Universal Robots URScript: FaiChun_9 Jan_Mcam1.script

def Machining1():
  # Default parameters:
  global speed_ms = 0.05
  global speed_rads = 0.75
  global accel_mss = 3
  global accel_radss = 1.2
  global blend_radius_m = 0.0003

  # Add subprograms here
  # Start of main program
  # Program generated by RoboDK v5.6.8 for UR10e on 13/01/2025 15:21:15
  # Using nominal kinematics.
  blend_radius_m = 0.0003
  speed_ms = 0.05
  # set_reference(p[0.340000, -0.055000, 0.001500, 0.000000, 0.000000, 0.000000])
  set_tcp(p[0.000000, 0.000000, 0.252000, 0.000000, 0.000000, 0.000000])
  # Show Tool
  movej([0.369740, -1.015857, -2.630541, -1.065992, 1.570796, 1.940536],accel_radss,speed_rads,0,blend_radius_m)
  movel([0.369740, -1.070501, -2.672301, -0.969586, 1.570796, 1.940536],accel_mss,speed_ms,0,blend_radius_m)
  #SetTool218
  #M_RunCode6
  #SetRPM107900
  #M_RunCode3
  speed_ms = 0.05
  movel([0.369740, -1.102928, -2.692299, -0.917162, 1.570796, 1.940536],accel_mss,speed_ms,0,blend_radius_m)
  speed_ms = 0.017
  movel([0.369740, -1.139169, -2.711618, -0.861603, 1.570796, 1.940536],accel_mss,speed_ms,0,blend_radius_m)
  speed_ms = 0.051
  movel([0.740413, -1.151810, -2.706369, -0.854210, 1.570796, 2.311209],accel_mss,speed_ms,0,blend_radius_m)
  movel([0.532956, -1.474706, -2.506843, -0.730840, 1.570796, 2.103752],accel_mss,speed_ms,0,blend_radius_m)
  movel([0.260506, -1.469805, -2.510970, -0.731614, 1.570796, 1.831302],accel_mss,speed_ms,0,blend_radius_m)
  movel([0.369740, -1.139169, -2.711618, -0.861603, 1.570796, 1.940536],accel_mss,speed_ms,0,blend_radius_m)
  speed_ms = 0.05
  movel([0.369740, -1.070501, -2.672301, -0.969586, 1.570796, 1.940536],accel_mss,speed_ms,0,blend_radius_m)
  speed_ms = 0.051
  movel([0.403329, -1.072947, -2.671379, -0.968064, 1.570796, 1.974125],accel_mss,speed_ms,0,blend_radius_m)
  movel([0.403329, -1.105379, -2.691338, -0.915672, 1.570796, 1.974125],accel_mss,speed_ms,0,blend_radius_m)
  speed_ms = 0.017
  movel([0.403329, -1.141610, -2.710617, -0.860163, 1.570796, 1.974125],accel_mss,speed_ms,0,blend_radius_m)
  speed_ms = 0.051
  movel([0.704795, -1.151689, -2.706421, -0.854280, 1.570796, 2.275591],accel_mss,speed_ms,0,blend_radius_m)
  movel([0.696497, -1.164526, -2.700927, -0.846935, 1.570796, 2.267294],accel_mss,speed_ms,0,blend_radius_m)
  movel([0.703914, -1.166306, -2.700152, -0.845930, 1.570796, 2.274710],accel_mss,speed_ms,0,blend_radius_m)
  movel([0.706062, -1.163020, -2.701581, -0.847789, 1.570796, 2.276858],accel_mss,speed_ms,0,blend_radius_m)
  movel([0.701176, -1.161829, -2.702095, -0.848464, 1.570796, 2.271972],accel_mss,speed_ms,0,blend_radius_m)
  movel([0.707357, -1.152320, -2.706154, -0.853914, 1.570796, 2.278154],accel_mss,speed_ms,0,blend_radius_m)
  movel([0.714620, -1.154134, -2.705387, -0.852868, 1.570796, 2.285416],accel_mss,speed_ms,0,blend_radius_m)
  movel([0.710409, -1.160546, -2.702649, -0.849195, 1.570796, 2.281205],accel_mss,speed_ms,0,blend_radius_m)
  movel([0.712930, -1.161189, -2.702372, -0.848829, 1.570796, 2.283727],accel_mss,speed_ms,0,blend_radius_m)
  movel([0.717151, -1.154792, -2.705108, -0.852489, 1.570796, 2.287947],accel_mss,speed_ms,0,blend_radius_m)
  movel([0.724331, -1.156706, -2.704294, -0.851389, 1.570796, 2.295128],accel_mss,speed_ms,0,blend_radius_m)
  movel([0.720088, -1.163073, -2.701558, -0.847759, 1.570796, 2.290884],accel_mss,speed_ms,0,blend_radius_m)
  movel([0.724885, -1.164384, -2.700989, -0.847016, 1.570796, 2.295682],accel_mss,speed_ms,0,blend_radius_m)
  movel([0.718665, -1.173659, -2.696916, -0.841814, 1.570796, 2.289462],accel_mss,speed_ms,0,blend_radius_m)
  movel([0.713893, -1.172379, -2.697484, -0.842526, 1.570796, 2.284689],accel_mss,speed_ms,0,blend_radius_m)
  movel([0.711746, -1.175609, -2.696048, -0.840731, 1.570796, 2.282542],accel_mss,speed_ms,0,blend_radius_m)
  movel([0.716510, -1.176879, -2.695481, -0.840029, 1.570796, 2.287306],accel_mss,speed_ms,0,blend_radius_m)
  movel([0.710435, -1.185964, -2.691373, -0.835052, 1.570796, 2.281231],accel_mss,speed_ms,0,blend_radius_m)
  movel([0.703407, -1.184139, -2.692206, -0.836045, 1.570796, 2.274203],accel_mss,speed_ms,0,blend_radius_m)
  movel([0.707472, -1.177990, -2.694983, -0.839416, 1.570796, 2.278268],accel_mss,speed_ms,0,blend_radius_m)
  movel([0.704985, -1.177355, -2.695268, -0.839766, 1.570796, 2.275781],accel_mss,speed_ms,0,blend_radius_m)
  movel([0.698841, -1.186688, -2.691042, -0.834659, 1.570796, 2.269637],accel_mss,speed_ms,0,blend_radius_m)
  movel([0.708330, -1.189119, -2.689926, -0.833344, 1.570796, 2.279126],accel_mss,speed_ms,0,blend_radius_m)
  movel([0.541731, -1.451056, -2.526411, -0.734922, 1.570796, 2.112528],accel_mss,speed_ms,0,blend_radius_m)
  movel([0.533908, -1.449838, -2.527395, -0.735156, 1.570796, 2.104704],accel_mss,speed_ms,0,blend_radius_m)
  movel([0.530407, -1.455837, -2.522525, -0.734027, 1.570796, 2.101203],accel_mss,speed_ms,0,blend_radius_m)
  movel([0.532431, -1.456143, -2.522276, -0.733971, 1.570796, 2.103227],accel_mss,speed_ms,0,blend_radius_m)
  movel([0.534734, -1.452207, -2.525478, -0.734704, 1.570796, 2.105531],accel_mss,speed_ms,0,blend_radius_m)
  movel([0.540507, -1.453110, -2.524746, -0.734533, 1.570796, 2.111303],accel_mss,speed_ms,0,blend_radius_m)
  movel([0.537071, -1.458916, -2.520004, -0.733469, 1.570796, 2.107867],accel_mss,speed_ms,0,blend_radius_m)
  movel([0.533196, -1.458312, -2.520500, -0.733577, 1.570796, 2.103992],accel_mss,speed_ms,0,blend_radius_m)
  movel([0.532009, -1.460340, -2.518833, -0.733216, 1.570796, 2.102805],accel_mss,speed_ms,0,blend_radius_m)
  movel([0.535879, -1.460941, -2.518338, -0.733110, 1.570796, 2.106675],accel_mss,speed_ms,0,blend_radius_m)
  movel([0.532503, -1.466680, -2.513581, -0.732128, 1.570796, 2.103300],accel_mss,speed_ms,0,blend_radius_m)
  movel([0.528655, -1.466088, -2.514074, -0.732226, 1.570796, 2.099451],accel_mss,speed_ms,0,blend_radius_m)
  movel([0.526411, -1.469942, -2.510855, -0.731592, 1.570796, 2.097208],accel_mss,speed_ms,0,blend_radius_m)
  movel([0.520712, -1.469102, -2.511559, -0.731728, 1.570796, 2.091509],accel_mss,speed_ms,0,blend_radius_m)
  movel([0.522933, -1.465238, -2.514782, -0.732370, 1.570796, 2.093730],accel_mss,speed_ms,0,blend_radius_m)
  movel([0.520922, -1.464950, -2.515020, -0.732418, 1.570796, 2.091718],accel_mss,speed_ms,0,blend_radius_m)
  movel([0.518707, -1.468815, -2.511798, -0.731775, 1.570796, 2.089503],accel_mss,speed_ms,0,blend_radius_m)
  movel([0.512973, -1.468021, -2.512463, -0.731905, 1.570796, 2.083769],accel_mss,speed_ms,0,blend_radius_m)
  movel([0.516230, -1.462277, -2.517236, -0.732877, 1.570796, 2.087027],accel_mss,speed_ms,0,blend_radius_m)
  movel([0.520125, -1.462817, -2.516788, -0.732783, 1.570796, 2.090921],accel_mss,speed_ms,0,blend_radius_m)
  movel([0.521283, -1.460796, -2.518457, -0.733135, 1.570796, 2.092080],accel_mss,speed_ms,0,blend_radius_m)
  movel([0.515352, -1.459974, -2.519134, -0.733281, 1.570796, 2.086148],accel_mss,speed_ms,0,blend_radius_m)
  movel([0.510955, -1.467752, -2.512687, -0.731950, 1.570796, 2.081751],accel_mss,speed_ms,0,blend_radius_m)
  movel([0.287607, -1.463384, -2.516319, -0.732685, 1.570796, 1.858403],accel_mss,speed_ms,0,blend_radius_m)
  movel([0.290165, -1.455515, -2.522788, -0.734086, 1.570796, 1.860961],accel_mss,speed_ms,0,blend_radius_m)
  movel([0.283577, -1.456094, -2.522316, -0.733980, 1.570796, 1.854374],accel_mss,speed_ms,0,blend_radius_m)
  movel([0.282922, -1.458141, -2.520640, -0.733608, 1.570796, 1.853718],accel_mss,speed_ms,0,blend_radius_m)
  movel([0.287251, -1.457756, -2.520955, -0.733677, 1.570796, 1.858048],accel_mss,speed_ms,0,blend_radius_m)
  movel([0.285369, -1.463569, -2.516166, -0.732654, 1.570796, 1.856165],accel_mss,speed_ms,0,blend_radius_m)
  movel([0.279002, -1.464133, -2.515698, -0.732557, 1.570796, 1.849799],accel_mss,speed_ms,0,blend_radius_m)
  movel([0.280240, -1.460222, -2.518931, -0.733237, 1.570796, 1.851036],accel_mss,speed_ms,0,blend_radius_m)
  movel([0.277998, -1.460430, -2.518759, -0.733200, 1.570796, 1.848794],accel_mss,speed_ms,0,blend_radius_m)
  movel([0.276770, -1.464340, -2.515527, -0.732522, 1.570796, 1.847566],accel_mss,speed_ms,0,blend_radius_m)
  movel([0.270394, -1.464949, -2.515021, -0.732418, 1.570796, 1.841191],accel_mss,speed_ms,0,blend_radius_m)
  movel([0.271594, -1.461046, -2.518252, -0.733092, 1.570796, 1.842390],accel_mss,speed_ms,0,blend_radius_m)
  movel([0.267266, -1.461483, -2.517891, -0.733015, 1.570796, 1.838062],accel_mss,speed_ms,0,blend_radius_m)
  movel([0.269033, -1.455666, -2.522665, -0.734058, 1.570796, 1.839830],accel_mss,speed_ms,0,blend_radius_m)
  movel([0.273388, -1.455222, -2.523027, -0.734140, 1.570796, 1.844184],accel_mss,speed_ms,0,blend_radius_m)
  movel([0.274023, -1.453169, -2.524697, -0.734522, 1.570796, 1.844820],accel_mss,speed_ms,0,blend_radius_m)
  movel([0.269656, -1.453615, -2.524335, -0.734439, 1.570796, 1.840452],accel_mss,speed_ms,0,blend_radius_m)
  movel([0.271457, -1.447728, -2.529094, -0.735567, 1.570796, 1.842253],accel_mss,speed_ms,0,blend_radius_m)
  movel([0.277970, -1.447061, -2.529630, -0.735698, 1.570796, 1.848766],accel_mss,speed_ms,0,blend_radius_m)
  movel([0.276719, -1.451051, -2.526415, -0.734923, 1.570796, 1.847516],accel_mss,speed_ms,0,blend_radius_m)
  movel([0.278991, -1.450829, -2.526594, -0.734966, 1.570796, 1.849787],accel_mss,speed_ms,0,blend_radius_m)
  movel([0.280907, -1.444757, -2.531476, -0.736156, 1.570796, 1.851704],accel_mss,speed_ms,0,blend_radius_m)
  movel([0.272096, -1.445651, -2.530761, -0.735977, 1.570796, 1.842893],accel_mss,speed_ms,0,blend_radius_m)
  movel([0.361539, -1.178261, -2.694862, -0.839266, 1.570796, 1.932335],accel_mss,speed_ms,0,blend_radius_m)
  movel([0.373305, -1.176443, -2.695676, -0.840270, 1.570796, 1.944101],accel_mss,speed_ms,0,blend_radius_m)
  movel([0.376834, -1.166854, -2.699913, -0.845622, 1.570796, 1.947630],accel_mss,speed_ms,0,blend_radius_m)
  movel([0.373758, -1.167323, -2.699708, -0.845358, 1.570796, 1.944554],accel_mss,speed_ms,0,blend_radius_m)
  movel([0.371445, -1.173642, -2.696924, -0.841824, 1.570796, 1.942241],accel_mss,speed_ms,0,blend_radius_m)
  movel([0.362714, -1.175005, -2.696318, -0.841066, 1.570796, 1.933510],accel_mss,speed_ms,0,blend_radius_m)
  movel([0.366061, -1.165657, -2.700435, -0.846297, 1.570796, 1.936857],accel_mss,speed_ms,0,blend_radius_m)
  movel([0.372018, -1.164705, -2.700850, -0.846834, 1.570796, 1.942815],accel_mss,speed_ms,0,blend_radius_m)
  movel([0.373227, -1.161386, -2.702286, -0.848716, 1.570796, 1.944024],accel_mss,speed_ms,0,blend_radius_m)
  movel([0.367253, -1.162346, -2.701872, -0.848171, 1.570796, 1.938049],accel_mss,speed_ms,0,blend_radius_m)
  movel([0.370690, -1.152795, -2.705954, -0.853640, 1.570796, 1.941486],accel_mss,speed_ms,0,blend_radius_m)
  movel([0.376724, -1.151811, -2.706369, -0.854209, 1.570796, 1.947521],accel_mss,speed_ms,0,blend_radius_m)
  movel([0.379122, -1.145259, -2.709109, -0.858021, 1.570796, 1.949918],accel_mss,speed_ms,0,blend_radius_m)
  movel([0.388102, -1.143842, -2.709696, -0.858851, 1.570796, 1.958898],accel_mss,speed_ms,0,blend_radius_m)
  movel([0.385643, -1.150419, -2.706955, -0.855015, 1.570796, 1.956439],accel_mss,speed_ms,0,blend_radius_m)
  movel([0.388764, -1.149949, -2.707152, -0.855288, 1.570796, 1.959560],accel_mss,speed_ms,0,blend_radius_m)
  movel([0.391247, -1.143361, -2.709895, -0.859133, 1.570796, 1.962043],accel_mss,speed_ms,0,blend_radius_m)
  movel([0.400196, -1.142054, -2.710434, -0.859901, 1.570796, 1.970993],accel_mss,speed_ms,0,blend_radius_m)
  movel([0.396453, -1.151808, -2.706370, -0.854211, 1.570796, 1.967249],accel_mss,speed_ms,0,blend_radius_m)
  movel([0.390466, -1.152664, -2.706009, -0.853716, 1.570796, 1.961262],accel_mss,speed_ms,0,blend_radius_m)
  movel([0.389190, -1.156041, -2.704577, -0.851771, 1.570796, 1.959986],accel_mss,speed_ms,0,blend_radius_m)
  movel([0.398252, -1.154767, -2.705119, -0.852504, 1.570796, 1.969048],accel_mss,speed_ms,0,blend_radius_m)
  movel([0.403329, -1.141610, -2.710617, -0.860163, 1.570796, 1.974125],accel_mss,speed_ms,0,blend_radius_m)
  speed_ms = 0.05
  movel([0.403329, -1.072947, -2.671379, -0.968064, 1.570796, 1.974125],accel_mss,speed_ms,0,blend_radius_m)
  #M_RunCode5
  speed_ms = 0.051
  movel([0.436039, -1.030309, -2.635411, -1.046670, 1.570796, 2.006835],accel_mss,speed_ms,0,blend_radius_m)
  #M_RunCode1
  #SetTool213
  #M_RunCode6
  #SetRPM107900
  #M_RunCode3
  speed_ms = 0.05
  movel([0.380621, -0.927251, -2.391546, -1.393592, 1.570796, 1.951417],accel_mss,speed_ms,0,blend_radius_m)
  speed_ms = 0.051
  movel([0.380621, -1.121069, -2.652122, -0.939198, 1.570796, 1.951417],accel_mss,speed_ms,0,blend_radius_m)
  movel([0.380621, -1.153481, -2.671325, -0.887584, 1.570796, 1.951417],accel_mss,speed_ms,0,blend_radius_m)
  speed_ms = 0.017
  movel([0.380621, -1.189377, -2.689807, -0.833205, 1.570796, 1.951417],accel_mss,speed_ms,0,blend_radius_m)
  speed_ms = 0.051
  movel([0.383999, -1.188172, -2.690361, -0.833856, 1.570796, 1.954796],accel_mss,speed_ms,0,blend_radius_m)
  movel([0.387929, -1.187302, -2.690760, -0.834326, 1.570796, 1.958725],accel_mss,speed_ms,0,blend_radius_m)
  movel([0.392921, -1.186724, -2.691025, -0.834640, 1.570796, 1.963717],accel_mss,speed_ms,0,blend_radius_m)
  movel([0.396406, -1.186468, -2.691143, -0.834778, 1.570796, 1.967202],accel_mss,speed_ms,0,blend_radius_m)
  movel([0.399894, -1.186176, -2.691276, -0.834937, 1.570796, 1.970690],accel_mss,speed_ms,0,blend_radius_m)
  movel([0.403055, -1.185763, -2.691465, -0.835161, 1.570796, 1.973851],accel_mss,speed_ms,0,blend_radius_m)
  movel([0.405472, -1.185291, -2.691681, -0.835418, 1.570796, 1.976268],accel_mss,speed_ms,0,blend_radius_m)
  movel([0.407571, -1.184727, -2.691938, -0.835724, 1.570796, 1.978367],accel_mss,speed_ms,0,blend_radius_m)
  movel([0.410903, -1.183473, -2.692508, -0.836408, 1.570796, 1.981699],accel_mss,speed_ms,0,blend_radius_m)
  movel([0.412588, -1.182637, -2.692888, -0.836864, 1.570796, 1.983384],accel_mss,speed_ms,0,blend_radius_m)
  movel([0.415576, -1.180774, -2.693730, -0.837884, 1.570796, 1.986373],accel_mss,speed_ms,0,blend_radius_m)
  movel([0.417237, -1.179418, -2.694342, -0.838629, 1.570796, 1.988033],accel_mss,speed_ms,0,blend_radius_m)
  movel([0.418646, -1.177700, -2.695113, -0.839575, 1.570796, 1.989443],accel_mss,speed_ms,0,blend_radius_m)
  movel([0.419750, -1.175666, -2.696023, -0.840700, 1.570796, 1.990546],accel_mss,speed_ms,0,blend_radius_m)
  movel([0.420402, -1.173479, -2.696996, -0.841914, 1.570796, 1.991198],accel_mss,speed_ms,0,blend_radius_m)
  movel([0.420438, -1.171501, -2.697872, -0.843016, 1.570796, 1.991235],accel_mss,speed_ms,0,blend_radius_m)
  movel([0.420217, -1.170743, -2.698207, -0.843440, 1.570796, 1.991013],accel_mss,speed_ms,0,blend_radius_m)
  movel([0.419855, -1.170173, -2.698457, -0.843759, 1.570796, 1.990652],accel_mss,speed_ms,0,blend_radius_m)
  movel([0.419383, -1.169789, -2.698626, -0.843973, 1.570796, 1.990180],accel_mss,speed_ms,0,blend_radius_m)
  movel([0.418119, -1.169559, -2.698728, -0.844102, 1.570796, 1.988915],accel_mss,speed_ms,0,blend_radius_m)
  movel([0.416505, -1.170034, -2.698519, -0.843836, 1.570796, 1.987302],accel_mss,speed_ms,0,blend_radius_m)
  movel([0.416237, -1.170163, -2.698462, -0.843764, 1.570796, 1.987034],accel_mss,speed_ms,0,blend_radius_m)
  movel([0.414985, -1.171929, -2.697683, -0.842778, 1.570796, 1.985782],accel_mss,speed_ms,0,blend_radius_m)
  movel([0.413492, -1.173744, -2.696878, -0.841766, 1.570796, 1.984288],accel_mss,speed_ms,0,blend_radius_m)
  movel([0.412436, -1.174807, -2.696406, -0.841176, 1.570796, 1.983232],accel_mss,speed_ms,0,blend_radius_m)
  movel([0.411578, -1.175521, -2.696088, -0.840780, 1.570796, 1.982374],accel_mss,speed_ms,0,blend_radius_m)
  movel([0.410708, -1.176097, -2.695830, -0.840461, 1.570796, 1.981504],accel_mss,speed_ms,0,blend_radius_m)
  movel([0.409905, -1.176478, -2.695660, -0.840250, 1.570796, 1.980701],accel_mss,speed_ms,0,blend_radius_m)
  movel([0.408376, -1.176754, -2.695537, -0.840098, 1.570796, 1.979172],accel_mss,speed_ms,0,blend_radius_m)
  movel([0.408234, -1.176742, -2.695542, -0.840104, 1.570796, 1.979030],accel_mss,speed_ms,0,blend_radius_m)
  movel([0.406466, -1.176296, -2.695742, -0.840351, 1.570796, 1.977262],accel_mss,speed_ms,0,blend_radius_m)
  movel([0.405390, -1.175348, -2.696165, -0.840876, 1.570796, 1.976186],accel_mss,speed_ms,0,blend_radius_m)
  movel([0.404939, -1.173986, -2.696771, -0.841632, 1.570796, 1.975735],accel_mss,speed_ms,0,blend_radius_m)
  movel([0.405099, -1.172279, -2.697528, -0.842582, 1.570796, 1.975896],accel_mss,speed_ms,0,blend_radius_m)
  movel([0.405880, -1.170338, -2.698385, -0.843666, 1.570796, 1.976676],accel_mss,speed_ms,0,blend_radius_m)
  movel([0.407213, -1.168390, -2.699241, -0.844758, 1.570796, 1.978009],accel_mss,speed_ms,0,blend_radius_m)
  movel([0.408857, -1.166781, -2.699945, -0.845663, 1.570796, 1.979653],accel_mss,speed_ms,0,blend_radius_m)
  movel([0.410787, -1.165550, -2.700482, -0.846357, 1.570796, 1.981584],accel_mss,speed_ms,0,blend_radius_m)
  movel([0.412791, -1.164886, -2.700771, -0.846732, 1.570796, 1.983588],accel_mss,speed_ms,0,blend_radius_m)
  movel([0.414812, -1.164846, -2.700788, -0.846754, 1.570796, 1.985608],accel_mss,speed_ms,0,blend_radius_m)
  movel([0.415507, -1.164994, -2.700724, -0.846671, 1.570796, 1.986303],accel_mss,speed_ms,0,blend_radius_m)
  movel([0.417738, -1.165921, -2.700320, -0.846148, 1.570796, 1.988534],accel_mss,speed_ms,0,blend_radius_m)
  movel([0.419793, -1.167599, -2.699588, -0.845203, 1.570796, 1.990590],accel_mss,speed_ms,0,blend_radius_m)
  movel([0.421507, -1.170024, -2.698523, -0.843842, 1.570796, 1.992303],accel_mss,speed_ms,0,blend_radius_m)
  movel([0.422695, -1.173065, -2.697180, -0.842144, 1.570796, 1.993492],accel_mss,speed_ms,0,blend_radius_m)
  movel([0.423223, -1.176462, -2.695668, -0.840259, 1.570796, 1.994019],accel_mss,speed_ms,0,blend_radius_m)
  movel([0.423058, -1.179904, -2.694123, -0.838362, 1.570796, 1.993854],accel_mss,speed_ms,0,blend_radius_m)
  movel([0.422274, -1.183152, -2.692654, -0.836583, 1.570796, 1.993070],accel_mss,speed_ms,0,blend_radius_m)
  movel([0.420984, -1.186080, -2.691320, -0.834989, 1.570796, 1.991781],accel_mss,speed_ms,0,blend_radius_m)
  movel([0.419277, -1.188669, -2.690133, -0.833587, 1.570796, 1.990074],accel_mss,speed_ms,0,blend_radius_m)
  movel([0.417187, -1.190952, -2.689080, -0.832357, 1.570796, 1.987983],accel_mss,speed_ms,0,blend_radius_m)
  movel([0.414698, -1.192969, -2.688145, -0.831275, 1.570796, 1.985494],accel_mss,speed_ms,0,blend_radius_m)
  movel([0.411744, -1.194743, -2.687319, -0.830327, 1.570796, 1.982541],accel_mss,speed_ms,0,blend_radius_m)
  movel([0.409937, -1.195593, -2.686922, -0.829874, 1.570796, 1.980733],accel_mss,speed_ms,0,blend_radius_m)
  movel([0.406912, -1.196699, -2.686405, -0.829286, 1.570796, 1.977709],accel_mss,speed_ms,0,blend_radius_m)
  movel([0.403445, -1.197467, -2.686044, -0.828878, 1.570796, 1.974241],accel_mss,speed_ms,0,blend_radius_m)
  movel([0.398983, -1.197989, -2.685799, -0.828601, 1.570796, 1.969779],accel_mss,speed_ms,0,blend_radius_m)
  movel([0.396138, -1.198246, -2.685678, -0.828465, 1.570796, 1.966934],accel_mss,speed_ms,0,blend_radius_m)
  movel([0.393290, -1.198591, -2.685516, -0.828282, 1.570796, 1.964086],accel_mss,speed_ms,0,blend_radius_m)
  movel([0.390854, -1.199043, -2.685303, -0.828043, 1.570796, 1.961650],accel_mss,speed_ms,0,blend_radius_m)
  movel([0.388892, -1.199570, -2.685054, -0.827764, 1.570796, 1.959688],accel_mss,speed_ms,0,blend_radius_m)
  movel([0.387163, -1.200181, -2.684766, -0.827442, 1.570796, 1.957959],accel_mss,speed_ms,0,blend_radius_m)
  movel([0.384322, -1.201557, -2.684115, -0.826717, 1.570796, 1.955118],accel_mss,speed_ms,0,blend_radius_m)
  movel([0.381459, -1.203495, -2.683194, -0.825700, 1.570796, 1.952256],accel_mss,speed_ms,0,blend_radius_m)
  movel([0.381214, -1.203689, -2.683102, -0.825599, 1.570796, 1.952010],accel_mss,speed_ms,0,blend_radius_m)
  movel([0.382206, -1.205244, -2.682360, -0.824786, 1.570796, 1.953002],accel_mss,speed_ms,0,blend_radius_m)
  movel([0.383252, -1.206538, -2.681740, -0.824111, 1.570796, 1.954048],accel_mss,speed_ms,0,blend_radius_m)
  movel([0.384343, -1.207588, -2.681236, -0.823565, 1.570796, 1.955140],accel_mss,speed_ms,0,blend_radius_m)
  movel([0.385467, -1.208411, -2.680840, -0.823138, 1.570796, 1.956263],accel_mss,speed_ms,0,blend_radius_m)
  movel([0.386616, -1.209027, -2.680543, -0.822819, 1.570796, 1.957413],accel_mss,speed_ms,0,blend_radius_m)
  movel([0.389049, -1.209700, -2.680218, -0.822471, 1.570796, 1.959845],accel_mss,speed_ms,0,blend_radius_m)
  movel([0.391565, -1.209683, -2.680226, -0.822480, 1.570796, 1.962362],accel_mss,speed_ms,0,blend_radius_m)
  movel([0.394197, -1.209043, -2.680535, -0.822811, 1.570796, 1.964993],accel_mss,speed_ms,0,blend_radius_m)
  movel([0.397008, -1.207785, -2.681141, -0.823463, 1.570796, 1.967805],accel_mss,speed_ms,0,blend_radius_m)
  movel([0.398343, -1.207009, -2.681514, -0.823866, 1.570796, 1.969139],accel_mss,speed_ms,0,blend_radius_m)
  movel([0.387393, -1.216041, -2.677132, -0.819216, 1.570796, 1.958190],accel_mss,speed_ms,0,blend_radius_m)
  movel([0.373654, -1.194729, -2.687326, -0.830334, 1.570796, 1.944450],accel_mss,speed_ms,0,blend_radius_m)
  movel([0.373249, -1.194112, -2.687613, -0.830664, 1.570796, 1.944045],accel_mss,speed_ms,0,blend_radius_m)
  movel([0.375328, -1.192380, -2.688418, -0.831590, 1.570796, 1.946125],accel_mss,speed_ms,0,blend_radius_m)
  movel([0.377499, -1.190904, -2.689102, -0.832383, 1.570796, 1.948295],accel_mss,speed_ms,0,blend_radius_m)
  movel([0.380387, -1.189467, -2.689765, -0.833156, 1.570796, 1.951184],accel_mss,speed_ms,0,blend_radius_m)
  movel([0.380621, -1.189377, -2.689807, -0.833205, 1.570796, 1.951417],accel_mss,speed_ms,0,blend_radius_m)
  speed_ms = 0.05
  movel([0.380621, -1.131501, -2.658598, -0.922290, 1.570796, 1.951417],accel_mss,speed_ms,0,blend_radius_m)
  speed_ms = 0.051
  movel([0.380621, -1.121069, -2.652122, -0.939198, 1.570796, 1.951417],accel_mss,speed_ms,0,blend_radius_m)
  movel([0.436617, -1.136722, -2.645392, -0.930276, 1.570796, 2.007413],accel_mss,speed_ms,0,blend_radius_m)
  movel([0.436617, -1.169075, -2.664345, -0.878969, 1.570796, 2.007413],accel_mss,speed_ms,0,blend_radius_m)
  speed_ms = 0.017
  movel([0.436617, -1.204809, -2.682567, -0.825012, 1.570796, 2.007413],accel_mss,speed_ms,0,blend_radius_m)
  speed_ms = 0.051
  movel([0.436929, -1.201228, -2.684271, -0.826890, 1.570796, 2.007725],accel_mss,speed_ms,0,blend_radius_m)
  movel([0.436607, -1.198383, -2.685614, -0.828392, 1.570796, 2.007404],accel_mss,speed_ms,0,blend_radius_m)
  movel([0.435725, -1.196201, -2.686638, -0.829550, 1.570796, 2.006521],accel_mss,speed_ms,0,blend_radius_m)
  movel([0.434327, -1.194619, -2.687377, -0.830393, 1.570796, 2.005124],accel_mss,speed_ms,0,blend_radius_m)
  movel([0.432439, -1.193606, -2.687849, -0.830934, 1.570796, 2.003236],accel_mss,speed_ms,0,blend_radius_m)
  movel([0.430057, -1.193161, -2.688056, -0.831172, 1.570796, 2.000854],accel_mss,speed_ms,0,blend_radius_m)
  movel([0.427169, -1.193310, -2.687987, -0.831093, 1.570796, 1.997965],accel_mss,speed_ms,0,blend_radius_m)
  movel([0.423785, -1.194095, -2.687621, -0.830673, 1.570796, 1.994581],accel_mss,speed_ms,0,blend_radius_m)
  movel([0.419952, -1.195561, -2.686937, -0.829891, 1.570796, 1.990748],accel_mss,speed_ms,0,blend_radius_m)
  movel([0.415791, -1.197705, -2.685933, -0.828752, 1.570796, 1.986587],accel_mss,speed_ms,0,blend_radius_m)
  movel([0.411494, -1.200472, -2.684628, -0.827289, 1.570796, 1.982291],accel_mss,speed_ms,0,blend_radius_m)
  movel([0.407314, -1.203723, -2.683086, -0.825581, 1.570796, 1.978110],accel_mss,speed_ms,0,blend_radius_m)
  movel([0.403492, -1.207275, -2.681386, -0.823728, 1.570796, 1.974289],accel_mss,speed_ms,0,blend_radius_m)
  movel([0.400216, -1.210938, -2.679619, -0.821832, 1.570796, 1.971012],accel_mss,speed_ms,0,blend_radius_m)
  movel([0.397587, -1.214561, -2.677856, -0.819971, 1.570796, 1.968383],accel_mss,speed_ms,0,blend_radius_m)
  movel([0.395632, -1.218046, -2.676147, -0.818196, 1.570796, 1.966428],accel_mss,speed_ms,0,blend_radius_m)
  movel([0.394335, -1.221348, -2.674514, -0.816526, 1.570796, 1.965132],accel_mss,speed_ms,0,blend_radius_m)
  movel([0.393990, -1.222635, -2.673875, -0.815879, 1.570796, 1.964786],accel_mss,speed_ms,0,blend_radius_m)
  movel([0.393819, -1.224825, -2.672782, -0.814782, 1.570796, 1.964615],accel_mss,speed_ms,0,blend_radius_m)
  movel([0.394040, -1.227752, -2.671313, -0.813324, 1.570796, 1.964836],accel_mss,speed_ms,0,blend_radius_m)
  movel([0.394806, -1.230002, -2.670177, -0.812210, 1.570796, 1.965602],accel_mss,speed_ms,0,blend_radius_m)
  movel([0.396055, -1.231651, -2.669341, -0.811398, 1.570796, 1.966851],accel_mss,speed_ms,0,blend_radius_m)
  movel([0.397753, -1.232760, -2.668776, -0.810853, 1.570796, 1.968549],accel_mss,speed_ms,0,blend_radius_m)
  movel([0.399903, -1.233347, -2.668477, -0.810565, 1.570796, 1.970700],accel_mss,speed_ms,0,blend_radius_m)
  movel([0.402512, -1.233403, -2.668448, -0.810537, 1.570796, 1.973308],accel_mss,speed_ms,0,blend_radius_m)
  movel([0.405590, -1.232897, -2.668707, -0.810786, 1.570796, 1.976387],accel_mss,speed_ms,0,blend_radius_m)
  movel([0.409117, -1.231781, -2.669274, -0.811333, 1.570796, 1.979913],accel_mss,speed_ms,0,blend_radius_m)
  movel([0.413019, -1.230039, -2.670158, -0.812192, 1.570796, 1.983815],accel_mss,speed_ms,0,blend_radius_m)
  movel([0.417152, -1.227681, -2.671349, -0.813359, 1.570796, 1.987948],accel_mss,speed_ms,0,blend_radius_m)
  movel([0.421305, -1.224793, -2.672798, -0.814798, 1.570796, 1.992102],accel_mss,speed_ms,0,blend_radius_m)
  movel([0.425243, -1.221512, -2.674433, -0.816444, 1.570796, 1.996040],accel_mss,speed_ms,0,blend_radius_m)
  movel([0.428757, -1.218010, -2.676165, -0.818214, 1.570796, 1.999553],accel_mss,speed_ms,0,blend_radius_m)
  movel([0.431708, -1.214438, -2.677916, -0.820034, 1.570796, 2.002504],accel_mss,speed_ms,0,blend_radius_m)
  movel([0.434028, -1.210915, -2.679630, -0.821844, 1.570796, 2.004824],accel_mss,speed_ms,0,blend_radius_m)
  movel([0.435711, -1.207501, -2.681278, -0.823610, 1.570796, 2.006508],accel_mss,speed_ms,0,blend_radius_m)
  movel([0.436617, -1.204809, -2.682567, -0.825012, 1.570796, 2.007413],accel_mss,speed_ms,0,blend_radius_m)
  speed_ms = 0.05
  movel([0.436617, -1.147144, -2.651786, -0.913459, 1.570796, 2.007413],accel_mss,speed_ms,0,blend_radius_m)
  speed_ms = 0.051
  movel([0.436617, -1.136722, -2.645392, -0.930276, 1.570796, 2.007413],accel_mss,speed_ms,0,blend_radius_m)
  movel([0.402334, -1.160294, -2.634802, -0.917293, 1.570796, 1.973130],accel_mss,speed_ms,0,blend_radius_m)
  movel([0.402334, -1.192513, -2.653378, -0.866497, 1.570796, 1.973130],accel_mss,speed_ms,0,blend_radius_m)
  speed_ms = 0.017
  movel([0.402334, -1.227961, -2.671208, -0.813220, 1.570796, 1.973130],accel_mss,speed_ms,0,blend_radius_m)
  speed_ms = 0.051
  movel([0.399988, -1.229223, -2.670571, -0.812595, 1.570796, 1.970785],accel_mss,speed_ms,0,blend_radius_m)
  movel([0.398129, -1.229756, -2.670301, -0.812331, 1.570796, 1.968925],accel_mss,speed_ms,0,blend_radius_m)
  movel([0.396798, -1.229657, -2.670351, -0.812381, 1.570796, 1.967595],accel_mss,speed_ms,0,blend_radius_m)
  movel([0.396017, -1.229029, -2.670669, -0.812691, 1.570796, 1.966813],accel_mss,speed_ms,0,blend_radius_m)
  movel([0.395804, -1.227950, -2.671213, -0.813226, 1.570796, 1.966601],accel_mss,speed_ms,0,blend_radius_m)
  movel([0.396204, -1.226474, -2.671955, -0.813959, 1.570796, 1.967001],accel_mss,speed_ms,0,blend_radius_m)
  movel([0.397291, -1.224647, -2.672871, -0.814871, 1.570796, 1.968087],accel_mss,speed_ms,0,blend_radius_m)
  movel([0.399106, -1.222568, -2.673908, -0.815913, 1.570796, 1.969902],accel_mss,speed_ms,0,blend_radius_m)
  movel([0.406141, -1.216101, -2.677103, -0.819185, 1.570796, 1.976937],accel_mss,speed_ms,0,blend_radius_m)
  movel([0.410949, -1.211934, -2.679136, -0.821319, 1.570796, 1.981745],accel_mss,speed_ms,0,blend_radius_m)
  movel([0.415358, -1.208284, -2.680901, -0.823204, 1.570796, 1.986154],accel_mss,speed_ms,0,blend_radius_m)
  movel([0.419212, -1.205255, -2.682354, -0.824780, 1.570796, 1.990008],accel_mss,speed_ms,0,blend_radius_m)
  movel([0.422503, -1.202824, -2.683513, -0.826052, 1.570796, 1.993299],accel_mss,speed_ms,0,blend_radius_m)
  movel([0.425265, -1.200931, -2.684411, -0.827047, 1.570796, 1.996061],accel_mss,speed_ms,0,blend_radius_m)
  movel([0.427550, -1.199513, -2.685081, -0.827795, 1.570796, 1.998346],accel_mss,speed_ms,0,blend_radius_m)
  movel([0.429412, -1.198496, -2.685560, -0.828332, 1.570796, 2.000209],accel_mss,speed_ms,0,blend_radius_m)
  movel([0.430916, -1.197811, -2.685882, -0.828695, 1.570796, 2.001712],accel_mss,speed_ms,0,blend_radius_m)
  movel([0.432108, -1.197407, -2.686072, -0.828909, 1.570796, 2.002904],accel_mss,speed_ms,0,blend_radius_m)
  movel([0.433044, -1.197228, -2.686156, -0.829004, 1.570796, 2.003841],accel_mss,speed_ms,0,blend_radius_m)
  movel([0.433768, -1.197232, -2.686155, -0.829003, 1.570796, 2.004564],accel_mss,speed_ms,0,blend_radius_m)
  movel([0.434743, -1.197712, -2.685929, -0.828748, 1.570796, 2.005539],accel_mss,speed_ms,0,blend_radius_m)
  movel([0.434902, -1.197930, -2.685827, -0.828633, 1.570796, 2.005698],accel_mss,speed_ms,0,blend_radius_m)
  movel([0.435050, -1.198509, -2.685554, -0.828325, 1.570796, 2.005846],accel_mss,speed_ms,0,blend_radius_m)
  movel([0.434852, -1.199802, -2.684945, -0.827642, 1.570796, 2.005648],accel_mss,speed_ms,0,blend_radius_m)
  movel([0.434006, -1.201486, -2.684148, -0.826754, 1.570796, 2.004803],accel_mss,speed_ms,0,blend_radius_m)
  movel([0.432321, -1.203737, -2.683079, -0.825573, 1.570796, 2.003117],accel_mss,speed_ms,0,blend_radius_m)
  movel([0.429506, -1.206736, -2.681645, -0.824008, 1.570796, 2.000303],accel_mss,speed_ms,0,blend_radius_m)
  movel([0.425244, -1.210649, -2.679759, -0.821981, 1.570796, 1.996041],accel_mss,speed_ms,0,blend_radius_m)
  movel([0.419297, -1.215560, -2.677368, -0.819461, 1.570796, 1.990093],accel_mss,speed_ms,0,blend_radius_m)
  movel([0.411783, -1.221286, -2.674545, -0.816558, 1.570796, 1.982579],accel_mss,speed_ms,0,blend_radius_m)
  movel([0.404088, -1.226777, -2.671803, -0.813809, 1.570796, 1.974885],accel_mss,speed_ms,0,blend_radius_m)
  movel([0.402334, -1.227961, -2.671208, -0.813220, 1.570796, 1.973130],accel_mss,speed_ms,0,blend_radius_m)
  speed_ms = 0.05
  movel([0.402334, -1.170687, -2.641073, -0.900629, 1.570796, 1.973130],accel_mss,speed_ms,0,blend_radius_m)
  speed_ms = 0.051
  movel([0.402334, -1.160294, -2.634802, -0.917293, 1.570796, 1.973130],accel_mss,speed_ms,0,blend_radius_m)
  movel([0.501584, -1.224318, -2.603129, -0.884943, 1.570796, 2.072381],accel_mss,speed_ms,0,blend_radius_m)
  movel([0.501584, -1.255923, -2.620674, -0.835791, 1.570796, 2.072381],accel_mss,speed_ms,0,blend_radius_m)
  speed_ms = 0.017
  movel([0.501584, -1.290346, -2.637441, -0.784602, 1.570796, 2.072381],accel_mss,speed_ms,0,blend_radius_m)
  speed_ms = 0.051
  movel([0.494290, -1.293714, -2.635480, -0.783195, 1.570796, 2.065087],accel_mss,speed_ms,0,blend_radius_m)
  movel([0.485005, -1.297578, -2.633213, -0.781598, 1.570796, 2.055802],accel_mss,speed_ms,0,blend_radius_m)
  movel([0.473858, -1.301828, -2.630697, -0.779864, 1.570796, 2.044654],accel_mss,speed_ms,0,blend_radius_m)
  movel([0.461472, -1.306187, -2.628092, -0.778111, 1.570796, 2.032268],accel_mss,speed_ms,0,blend_radius_m)
  movel([0.449108, -1.310193, -2.625675, -0.776520, 1.570796, 2.019904],accel_mss,speed_ms,0,blend_radius_m)
  movel([0.438420, -1.313296, -2.623790, -0.775304, 1.570796, 2.009216],accel_mss,speed_ms,0,blend_radius_m)
  movel([0.436376, -1.313832, -2.623462, -0.775095, 1.570796, 2.007172],accel_mss,speed_ms,0,blend_radius_m)
  movel([0.433761, -1.315367, -2.622523, -0.774498, 1.570796, 2.004557],accel_mss,speed_ms,0,blend_radius_m)
  movel([0.427766, -1.319278, -2.620117, -0.772994, 1.570796, 1.998563],accel_mss,speed_ms,0,blend_radius_m)
  movel([0.418182, -1.326018, -2.615923, -0.770449, 1.570796, 1.988978],accel_mss,speed_ms,0,blend_radius_m)
  movel([0.399906, -1.339314, -2.607467, -0.765608, 1.570796, 1.970702],accel_mss,speed_ms,0,blend_radius_m)
  movel([0.390441, -1.346141, -2.603032, -0.763217, 1.570796, 1.961238],accel_mss,speed_ms,0,blend_radius_m)
  movel([0.383665, -1.350921, -2.599887, -0.761581, 1.570796, 1.954462],accel_mss,speed_ms,0,blend_radius_m)
  movel([0.377983, -1.354824, -2.597296, -0.760269, 1.570796, 1.948779],accel_mss,speed_ms,0,blend_radius_m)
  movel([0.373032, -1.358117, -2.595093, -0.759178, 1.570796, 1.943829],accel_mss,speed_ms,0,blend_radius_m)
  movel([0.368648, -1.360925, -2.593203, -0.758261, 1.570796, 1.939445],accel_mss,speed_ms,0,blend_radius_m)
  movel([0.364735, -1.363325, -2.591579, -0.757485, 1.570796, 1.935531],accel_mss,speed_ms,0,blend_radius_m)
  movel([0.361224, -1.365372, -2.590187, -0.756830, 1.570796, 1.932020],accel_mss,speed_ms,0,blend_radius_m)
  movel([0.358064, -1.367110, -2.589000, -0.756279, 1.570796, 1.928860],accel_mss,speed_ms,0,blend_radius_m)
  movel([0.355217, -1.368570, -2.588001, -0.755819, 1.570796, 1.926013],accel_mss,speed_ms,0,blend_radius_m)
  movel([0.352648, -1.369782, -2.587168, -0.755439, 1.570796, 1.923444],accel_mss,speed_ms,0,blend_radius_m)
  movel([0.350331, -1.370771, -2.586487, -0.755131, 1.570796, 1.921127],accel_mss,speed_ms,0,blend_radius_m)
  movel([0.348238, -1.371561, -2.585942, -0.754886, 1.570796, 1.919034],accel_mss,speed_ms,0,blend_radius_m)
  movel([0.346349, -1.372171, -2.585521, -0.754697, 1.570796, 1.917145],accel_mss,speed_ms,0,blend_radius_m)
  movel([0.343034, -1.372927, -2.584998, -0.754464, 1.570796, 1.913830],accel_mss,speed_ms,0,blend_radius_m)
  movel([0.340352, -1.373115, -2.584868, -0.754406, 1.570796, 1.911149],accel_mss,speed_ms,0,blend_radius_m)
  movel([0.338182, -1.372819, -2.585072, -0.754497, 1.570796, 1.908978],accel_mss,speed_ms,0,blend_radius_m)
  movel([0.336427, -1.372082, -2.585582, -0.754725, 1.570796, 1.907224],accel_mss,speed_ms,0,blend_radius_m)
  movel([0.335034, -1.370899, -2.586399, -0.755091, 1.570796, 1.905830],accel_mss,speed_ms,0,blend_radius_m)
  movel([0.333980, -1.369226, -2.587550, -0.755613, 1.570796, 1.904777],accel_mss,speed_ms,0,blend_radius_m)
  movel([0.333279, -1.366978, -2.589091, -0.756320, 1.570796, 1.904075],accel_mss,speed_ms,0,blend_radius_m)
  movel([0.332983, -1.364041, -2.591093, -0.757255, 1.570796, 1.903780],accel_mss,speed_ms,0,blend_radius_m)
  movel([0.333172, -1.360271, -2.593644, -0.758473, 1.570796, 1.903968],accel_mss,speed_ms,0,blend_radius_m)
  movel([0.333950, -1.355498, -2.596847, -0.760044, 1.570796, 1.904746],accel_mss,speed_ms,0,blend_radius_m)
  movel([0.334305, -1.353900, -2.597912, -0.760577, 1.570796, 1.905101],accel_mss,speed_ms,0,blend_radius_m)
  movel([0.337015, -1.354939, -2.597219, -0.760230, 1.570796, 1.907812],accel_mss,speed_ms,0,blend_radius_m)
  movel([0.338299, -1.355337, -2.596954, -0.760098, 1.570796, 1.909096],accel_mss,speed_ms,0,blend_radius_m)
  movel([0.339090, -1.355435, -2.596889, -0.760065, 1.570796, 1.909886],accel_mss,speed_ms,0,blend_radius_m)
  movel([0.339937, -1.355391, -2.596918, -0.760080, 1.570796, 1.910733],accel_mss,speed_ms,0,blend_radius_m)
  movel([0.341287, -1.355001, -2.597178, -0.760210, 1.570796, 1.912083],accel_mss,speed_ms,0,blend_radius_m)
  movel([0.343418, -1.353946, -2.597881, -0.760562, 1.570796, 1.914215],accel_mss,speed_ms,0,blend_radius_m)
  movel([0.346600, -1.351932, -2.599218, -0.761239, 1.570796, 1.917397],accel_mss,speed_ms,0,blend_radius_m)
  movel([0.351189, -1.348589, -2.601425, -0.762375, 1.570796, 1.921985],accel_mss,speed_ms,0,blend_radius_m)
  movel([0.357580, -1.343508, -2.604750, -0.764131, 1.570796, 1.928376],accel_mss,speed_ms,0,blend_radius_m)
  movel([0.366212, -1.336274, -2.609422, -0.766694, 1.570796, 1.937008],accel_mss,speed_ms,0,blend_radius_m)
  movel([0.376307, -1.327749, -2.614835, -0.769805, 1.570796, 1.947103],accel_mss,speed_ms,0,blend_radius_m)
  movel([0.390474, -1.317109, -2.621454, -0.773826, 1.570796, 1.961271],accel_mss,speed_ms,0,blend_radius_m)
  movel([0.383241, -1.318954, -2.620317, -0.773118, 1.570796, 1.954037],accel_mss,speed_ms,0,blend_radius_m)
  movel([0.375997, -1.320426, -2.619407, -0.772556, 1.570796, 1.946793],accel_mss,speed_ms,0,blend_radius_m)
  movel([0.369750, -1.321281, -2.618877, -0.772231, 1.570796, 1.940547],accel_mss,speed_ms,0,blend_radius_m)
  movel([0.364410, -1.321585, -2.618688, -0.772116, 1.570796, 1.935206],accel_mss,speed_ms,0,blend_radius_m)
  movel([0.359884, -1.321397, -2.618805, -0.772187, 1.570796, 1.930680],accel_mss,speed_ms,0,blend_radius_m)
  movel([0.356095, -1.320765, -2.619197, -0.772427, 1.570796, 1.926891],accel_mss,speed_ms,0,blend_radius_m)
  movel([0.352970, -1.319736, -2.619834, -0.772819, 1.570796, 1.923767],accel_mss,speed_ms,0,blend_radius_m)
  movel([0.350449, -1.318334, -2.620700, -0.773355, 1.570796, 1.921246],accel_mss,speed_ms,0,blend_radius_m)
  movel([0.348482, -1.316585, -2.621776, -0.774028, 1.570796, 1.919278],accel_mss,speed_ms,0,blend_radius_m)
  movel([0.347038, -1.314497, -2.623056, -0.774836, 1.570796, 1.917835],accel_mss,speed_ms,0,blend_radius_m)
  movel([0.346099, -1.312064, -2.624539, -0.775785, 1.570796, 1.916895],accel_mss,speed_ms,0,blend_radius_m)
  movel([0.345661, -1.309283, -2.626226, -0.776880, 1.570796, 1.916457],accel_mss,speed_ms,0,blend_radius_m)
  movel([0.345745, -1.306140, -2.628119, -0.778129, 1.570796, 1.916542],accel_mss,speed_ms,0,blend_radius_m)
  movel([0.346374, -1.302637, -2.630215, -0.779537, 1.570796, 1.917171],accel_mss,speed_ms,0,blend_radius_m)
  movel([0.347579, -1.298790, -2.632498, -0.781101, 1.570796, 1.918375],accel_mss,speed_ms,0,blend_radius_m)
  movel([0.349372, -1.294658, -2.634928, -0.782803, 1.570796, 1.920168],accel_mss,speed_ms,0,blend_radius_m)
  movel([0.351743, -1.290340, -2.637444, -0.784605, 1.570796, 1.922539],accel_mss,speed_ms,0,blend_radius_m)
  movel([0.354623, -1.286008, -2.639945, -0.786436, 1.570796, 1.925419],accel_mss,speed_ms,0,blend_radius_m)
  movel([0.357881, -1.281879, -2.642305, -0.788205, 1.570796, 1.928677],accel_mss,speed_ms,0,blend_radius_m)
  movel([0.361327, -1.278187, -2.644398, -0.789804, 1.570796, 1.932123],accel_mss,speed_ms,0,blend_radius_m)
  movel([0.364750, -1.275125, -2.646121, -0.791143, 1.570796, 1.935546],accel_mss,speed_ms,0,blend_radius_m)
  movel([0.367969, -1.272801, -2.647421, -0.792167, 1.570796, 1.938766],accel_mss,speed_ms,0,blend_radius_m)
  movel([0.370877, -1.271219, -2.648301, -0.792869, 1.570796, 1.941673],accel_mss,speed_ms,0,blend_radius_m)
  movel([0.373430, -1.270330, -2.648795, -0.793264, 1.570796, 1.944227],accel_mss,speed_ms,0,blend_radius_m)
  movel([0.375649, -1.270060, -2.648945, -0.793384, 1.570796, 1.946445],accel_mss,speed_ms,0,blend_radius_m)
  movel([0.377564, -1.270368, -2.648774, -0.793247, 1.570796, 1.948360],accel_mss,speed_ms,0,blend_radius_m)
  movel([0.378012, -1.270541, -2.648678, -0.793170, 1.570796, 1.948809],accel_mss,speed_ms,0,blend_radius_m)
  movel([0.375550, -1.271287, -2.648264, -0.792838, 1.570796, 1.946347],accel_mss,speed_ms,0,blend_radius_m)
  movel([0.372751, -1.272532, -2.647570, -0.792286, 1.570796, 1.943548],accel_mss,speed_ms,0,blend_radius_m)
  movel([0.370655, -1.273915, -2.646799, -0.791676, 1.570796, 1.941451],accel_mss,speed_ms,0,blend_radius_m)
  movel([0.369146, -1.275381, -2.645978, -0.791031, 1.570796, 1.939942],accel_mss,speed_ms,0,blend_radius_m)
  movel([0.368128, -1.276919, -2.645113, -0.790357, 1.570796, 1.938924],accel_mss,speed_ms,0,blend_radius_m)
  movel([0.367564, -1.278548, -2.644194, -0.789646, 1.570796, 1.938360],accel_mss,speed_ms,0,blend_radius_m)
  movel([0.367478, -1.280272, -2.643218, -0.788898, 1.570796, 1.938275],accel_mss,speed_ms,0,blend_radius_m)
  movel([0.367952, -1.282053, -2.642206, -0.788129, 1.570796, 1.938748],accel_mss,speed_ms,0,blend_radius_m)
  movel([0.369064, -1.283784, -2.641219, -0.787386, 1.570796, 1.939860],accel_mss,speed_ms,0,blend_radius_m)
  movel([0.370834, -1.285299, -2.640351, -0.786738, 1.570796, 1.941630],accel_mss,speed_ms,0,blend_radius_m)
  movel([0.373185, -1.286430, -2.639702, -0.786257, 1.570796, 1.943981],accel_mss,speed_ms,0,blend_radius_m)
  movel([0.374119, -1.286713, -2.639539, -0.786137, 1.570796, 1.944915],accel_mss,speed_ms,0,blend_radius_m)
  movel([0.377254, -1.286882, -2.639442, -0.786065, 1.570796, 1.948050],accel_mss,speed_ms,0,blend_radius_m)
  movel([0.382371, -1.286683, -2.639556, -0.786149, 1.570796, 1.953168],accel_mss,speed_ms,0,blend_radius_m)
  movel([0.389141, -1.285937, -2.639985, -0.786467, 1.570796, 1.959937],accel_mss,speed_ms,0,blend_radius_m)
  movel([0.397793, -1.284542, -2.640785, -0.787062, 1.570796, 1.968590],accel_mss,speed_ms,0,blend_radius_m)
  movel([0.408447, -1.282431, -2.641991, -0.787967, 1.570796, 1.979243],accel_mss,speed_ms,0,blend_radius_m)
  movel([0.420958, -1.279597, -2.643601, -0.789191, 1.570796, 1.991754],accel_mss,speed_ms,0,blend_radius_m)
  movel([0.434586, -1.276199, -2.645518, -0.790672, 1.570796, 2.005383],accel_mss,speed_ms,0,blend_radius_m)
  movel([0.447369, -1.272713, -2.647470, -0.792206, 1.570796, 2.018165],accel_mss,speed_ms,0,blend_radius_m)
  movel([0.447557, -1.272657, -2.647501, -0.792231, 1.570796, 2.018353],accel_mss,speed_ms,0,blend_radius_m)
  movel([0.448346, -1.272216, -2.647747, -0.792426, 1.570796, 2.019142],accel_mss,speed_ms,0,blend_radius_m)
  movel([0.448612, -1.271950, -2.647895, -0.792544, 1.570796, 2.019408],accel_mss,speed_ms,0,blend_radius_m)
  movel([0.448671, -1.271485, -2.648153, -0.792750, 1.570796, 2.019467],accel_mss,speed_ms,0,blend_radius_m)
  movel([0.448335, -1.270925, -2.648465, -0.792999, 1.570796, 2.019132],accel_mss,speed_ms,0,blend_radius_m)
  movel([0.447403, -1.269942, -2.649010, -0.793437, 1.570796, 2.018199],accel_mss,speed_ms,0,blend_radius_m)
  movel([0.445446, -1.268639, -2.649731, -0.794019, 1.570796, 2.016242],accel_mss,speed_ms,0,blend_radius_m)
  movel([0.442408, -1.267319, -2.650459, -0.794610, 1.570796, 2.013204],accel_mss,speed_ms,0,blend_radius_m)
  movel([0.438040, -1.265514, -2.651452, -0.795423, 1.570796, 2.008836],accel_mss,speed_ms,0,blend_radius_m)
  movel([0.436430, -1.264616, -2.651944, -0.795829, 1.570796, 2.007227],accel_mss,speed_ms,0,blend_radius_m)
  movel([0.435166, -1.263706, -2.652442, -0.796241, 1.570796, 2.005963],accel_mss,speed_ms,0,blend_radius_m)
  movel([0.434122, -1.262734, -2.652973, -0.796682, 1.570796, 2.004918],accel_mss,speed_ms,0,blend_radius_m)
  movel([0.433245, -1.261679, -2.653547, -0.797162, 1.570796, 2.004041],accel_mss,speed_ms,0,blend_radius_m)
  movel([0.431906, -1.259192, -2.654897, -0.798300, 1.570796, 2.002702],accel_mss,speed_ms,0,blend_radius_m)
  movel([0.431115, -1.256187, -2.656517, -0.799685, 1.570796, 2.001911],accel_mss,speed_ms,0,blend_radius_m)
  movel([0.430874, -1.252521, -2.658479, -0.801389, 1.570796, 2.001671],accel_mss,speed_ms,0,blend_radius_m)
  movel([0.430908, -1.251391, -2.659080, -0.801918, 1.570796, 2.001705],accel_mss,speed_ms,0,blend_radius_m)
  movel([0.430987, -1.249743, -2.659954, -0.802692, 1.570796, 2.001783],accel_mss,speed_ms,0,blend_radius_m)
  movel([0.431577, -1.246568, -2.661630, -0.804191, 1.570796, 2.002373],accel_mss,speed_ms,0,blend_radius_m)
  movel([0.432763, -1.243119, -2.663436, -0.805834, 1.570796, 2.003559],accel_mss,speed_ms,0,blend_radius_m)
  movel([0.434580, -1.239363, -2.665387, -0.807639, 1.570796, 2.005376],accel_mss,speed_ms,0,blend_radius_m)
  movel([0.437087, -1.235273, -2.667493, -0.809624, 1.570796, 2.007883],accel_mss,speed_ms,0,blend_radius_m)
  movel([0.440338, -1.230830, -2.669757, -0.811802, 1.570796, 2.011134],accel_mss,speed_ms,0,blend_radius_m)
  movel([0.444383, -1.226054, -2.672166, -0.814168, 1.570796, 2.015179],accel_mss,speed_ms,0,blend_radius_m)
  movel([0.449224, -1.221012, -2.674681, -0.816696, 1.570796, 2.020020],accel_mss,speed_ms,0,blend_radius_m)
  movel([0.454785, -1.215845, -2.677228, -0.819316, 1.570796, 2.025581],accel_mss,speed_ms,0,blend_radius_m)
  movel([0.460857, -1.210792, -2.679690, -0.821907, 1.570796, 2.031654],accel_mss,speed_ms,0,blend_radius_m)
  movel([0.467052, -1.206211, -2.681897, -0.824281, 1.570796, 2.037848],accel_mss,speed_ms,0,blend_radius_m)
  movel([0.472819, -1.202492, -2.683671, -0.826226, 1.570796, 2.043615],accel_mss,speed_ms,0,blend_radius_m)
  movel([0.477386, -1.200045, -2.684830, -0.827514, 1.570796, 2.048183],accel_mss,speed_ms,0,blend_radius_m)
  movel([0.482593, -1.197853, -2.685863, -0.828673, 1.570796, 2.053389],accel_mss,speed_ms,0,blend_radius_m)
  movel([0.489106, -1.195587, -2.686925, -0.829877, 1.570796, 2.059903],accel_mss,speed_ms,0,blend_radius_m)
  movel([0.494832, -1.194146, -2.687597, -0.830645, 1.570796, 2.065628],accel_mss,speed_ms,0,blend_radius_m)
  movel([0.499874, -1.193446, -2.687923, -0.831020, 1.570796, 2.070671],accel_mss,speed_ms,0,blend_radius_m)
  movel([0.504327, -1.193410, -2.687940, -0.831039, 1.570796, 2.075124],accel_mss,speed_ms,0,blend_radius_m)
  movel([0.508280, -1.193996, -2.687667, -0.830726, 1.570796, 2.079076],accel_mss,speed_ms,0,blend_radius_m)
  movel([0.511809, -1.195188, -2.687111, -0.830089, 1.570796, 2.082605],accel_mss,speed_ms,0,blend_radius_m)
  movel([0.514990, -1.196997, -2.686265, -0.829127, 1.570796, 2.085786],accel_mss,speed_ms,0,blend_radius_m)
  movel([0.517899, -1.199486, -2.685094, -0.827809, 1.570796, 2.088695],accel_mss,speed_ms,0,blend_radius_m)
  movel([0.520641, -1.202774, -2.683537, -0.826078, 1.570796, 2.091437],accel_mss,speed_ms,0,blend_radius_m)
  movel([0.523434, -1.207190, -2.681427, -0.823772, 1.570796, 2.094230],accel_mss,speed_ms,0,blend_radius_m)
  movel([0.527325, -1.214218, -2.678024, -0.820147, 1.570796, 2.098121],accel_mss,speed_ms,0,blend_radius_m)
  movel([0.529065, -1.216981, -2.676671, -0.818737, 1.570796, 2.099862],accel_mss,speed_ms,0,blend_radius_m)
  movel([0.530481, -1.218857, -2.675747, -0.817785, 1.570796, 2.101277],accel_mss,speed_ms,0,blend_radius_m)
  movel([0.531812, -1.220310, -2.675029, -0.817050, 1.570796, 2.102608],accel_mss,speed_ms,0,blend_radius_m)
  movel([0.533127, -1.221465, -2.674456, -0.816467, 1.570796, 2.103924],accel_mss,speed_ms,0,blend_radius_m)
  movel([0.534457, -1.222390, -2.673997, -0.816002, 1.570796, 2.105253],accel_mss,speed_ms,0,blend_radius_m)
  movel([0.535819, -1.223114, -2.673636, -0.815639, 1.570796, 2.106615],accel_mss,speed_ms,0,blend_radius_m)
  movel([0.538758, -1.224063, -2.673163, -0.815163, 1.570796, 2.109554],accel_mss,speed_ms,0,blend_radius_m)
  movel([0.541977, -1.224372, -2.673008, -0.815008, 1.570796, 2.112773],accel_mss,speed_ms,0,blend_radius_m)
  movel([0.545580, -1.224079, -2.673155, -0.815155, 1.570796, 2.116376],accel_mss,speed_ms,0,blend_radius_m)
  movel([0.547123, -1.223793, -2.673298, -0.815298, 1.570796, 2.117920],accel_mss,speed_ms,0,blend_radius_m)
  movel([0.550189, -1.222807, -2.673790, -0.815793, 1.570796, 2.120985],accel_mss,speed_ms,0,blend_radius_m)
  movel([0.552790, -1.221470, -2.674454, -0.816465, 1.570796, 2.123586],accel_mss,speed_ms,0,blend_radius_m)
  movel([0.555070, -1.219805, -2.675279, -0.817305, 1.570796, 2.125866],accel_mss,speed_ms,0,blend_radius_m)
  movel([0.557046, -1.217835, -2.676251, -0.818303, 1.570796, 2.127842],accel_mss,speed_ms,0,blend_radius_m)
  movel([0.558707, -1.215585, -2.677356, -0.819449, 1.570796, 2.129503],accel_mss,speed_ms,0,blend_radius_m)
  movel([0.559993, -1.213101, -2.678569, -0.820720, 1.570796, 2.130789],accel_mss,speed_ms,0,blend_radius_m)
  movel([0.560815, -1.210500, -2.679831, -0.822058, 1.570796, 2.131612],accel_mss,speed_ms,0,blend_radius_m)
  movel([0.561069, -1.207979, -2.681048, -0.823362, 1.570796, 2.131866],accel_mss,speed_ms,0,blend_radius_m)
  movel([0.560702, -1.205792, -2.682098, -0.824500, 1.570796, 2.131499],accel_mss,speed_ms,0,blend_radius_m)
  movel([0.559745, -1.204154, -2.682880, -0.825355, 1.570796, 2.130541],accel_mss,speed_ms,0,blend_radius_m)
  movel([0.558294, -1.203166, -2.683351, -0.825872, 1.570796, 2.129090],accel_mss,speed_ms,0,blend_radius_m)
  movel([0.556438, -1.202838, -2.683506, -0.826044, 1.570796, 2.127235],accel_mss,speed_ms,0,blend_radius_m)
  movel([0.554213, -1.203162, -2.683353, -0.825875, 1.570796, 2.125009],accel_mss,speed_ms,0,blend_radius_m)
  movel([0.551613, -1.204161, -2.682877, -0.825352, 1.570796, 2.122409],accel_mss,speed_ms,0,blend_radius_m)
  movel([0.548596, -1.205908, -2.682042, -0.824439, 1.570796, 2.119392],accel_mss,speed_ms,0,blend_radius_m)
  movel([0.548413, -1.206030, -2.681983, -0.824375, 1.570796, 2.119209],accel_mss,speed_ms,0,blend_radius_m)
  movel([0.550095, -1.206356, -2.681827, -0.824206, 1.570796, 2.120891],accel_mss,speed_ms,0,blend_radius_m)
  movel([0.551454, -1.207197, -2.681423, -0.823768, 1.570796, 2.122251],accel_mss,speed_ms,0,blend_radius_m)
  movel([0.552060, -1.208385, -2.680852, -0.823152, 1.570796, 2.122856],accel_mss,speed_ms,0,blend_radius_m)
  movel([0.551991, -1.209795, -2.680172, -0.822422, 1.570796, 2.122788],accel_mss,speed_ms,0,blend_radius_m)
  movel([0.551305, -1.211367, -2.679411, -0.821611, 1.570796, 2.122102],accel_mss,speed_ms,0,blend_radius_m)
  movel([0.549987, -1.213082, -2.678578, -0.820729, 1.570796, 2.120783],accel_mss,speed_ms,0,blend_radius_m)
  movel([0.547965, -1.214919, -2.677682, -0.819789, 1.570796, 2.118762],accel_mss,speed_ms,0,blend_radius_m)
  movel([0.547458, -1.215305, -2.677492, -0.819591, 1.570796, 2.118254],accel_mss,speed_ms,0,blend_radius_m)
  movel([0.545627, -1.216551, -2.676882, -0.818956, 1.570796, 2.116423],accel_mss,speed_ms,0,blend_radius_m)
  movel([0.542919, -1.217967, -2.676186, -0.818236, 1.570796, 2.113716],accel_mss,speed_ms,0,blend_radius_m)
  movel([0.540409, -1.218777, -2.675787, -0.817825, 1.570796, 2.111205],accel_mss,speed_ms,0,blend_radius_m)
  movel([0.538072, -1.219014, -2.675670, -0.817705, 1.570796, 2.108868],accel_mss,speed_ms,0,blend_radius_m)
  movel([0.535895, -1.218681, -2.675834, -0.817874, 1.570796, 2.106691],accel_mss,speed_ms,0,blend_radius_m)
  movel([0.533905, -1.217741, -2.676297, -0.818351, 1.570796, 2.104702],accel_mss,speed_ms,0,blend_radius_m)
  movel([0.532160, -1.216153, -2.677077, -0.819159, 1.570796, 2.102957],accel_mss,speed_ms,0,blend_radius_m)
  movel([0.530763, -1.213899, -2.678180, -0.820310, 1.570796, 2.101560],accel_mss,speed_ms,0,blend_radius_m)
  movel([0.529830, -1.211022, -2.679578, -0.821789, 1.570796, 2.100627],accel_mss,speed_ms,0,blend_radius_m)
  movel([0.529472, -1.207644, -2.681209, -0.823536, 1.570796, 2.100268],accel_mss,speed_ms,0,blend_radius_m)
  movel([0.529745, -1.203955, -2.682975, -0.825459, 1.570796, 2.100541],accel_mss,speed_ms,0,blend_radius_m)
  movel([0.530636, -1.200167, -2.684773, -0.827450, 1.570796, 2.101433],accel_mss,speed_ms,0,blend_radius_m)
  movel([0.532101, -1.196443, -2.686524, -0.829421, 1.570796, 2.102897],accel_mss,speed_ms,0,blend_radius_m)
  movel([0.534065, -1.192902, -2.688176, -0.831311, 1.570796, 2.104861],accel_mss,speed_ms,0,blend_radius_m)
  movel([0.536476, -1.189590, -2.689709, -0.833090, 1.570796, 2.107273],accel_mss,speed_ms,0,blend_radius_m)
  movel([0.539304, -1.186530, -2.691114, -0.834745, 1.570796, 2.110101],accel_mss,speed_ms,0,blend_radius_m)
  movel([0.542551, -1.183720, -2.692396, -0.836273, 1.570796, 2.113348],accel_mss,speed_ms,0,blend_radius_m)
  movel([0.546240, -1.181174, -2.693550, -0.837665, 1.570796, 2.117036],accel_mss,speed_ms,0,blend_radius_m)
  movel([0.546537, -1.180990, -2.693633, -0.837766, 1.570796, 2.117334],accel_mss,speed_ms,0,blend_radius_m)
  movel([0.550942, -1.178476, -2.694765, -0.839148, 1.570796, 2.121738],accel_mss,speed_ms,0,blend_radius_m)
  movel([0.555378, -1.176501, -2.695650, -0.840238, 1.570796, 2.126174],accel_mss,speed_ms,0,blend_radius_m)
  movel([0.559795, -1.175103, -2.696274, -0.841012, 1.570796, 2.130592],accel_mss,speed_ms,0,blend_radius_m)
  movel([0.564115, -1.174313, -2.696626, -0.841450, 1.570796, 2.134911],accel_mss,speed_ms,0,blend_radius_m)
  movel([0.568237, -1.174165, -2.696691, -0.841532, 1.570796, 2.139034],accel_mss,speed_ms,0,blend_radius_m)
  movel([0.572053, -1.174678, -2.696463, -0.841248, 1.570796, 2.142849],accel_mss,speed_ms,0,blend_radius_m)
  movel([0.575441, -1.175837, -2.695947, -0.840605, 1.570796, 2.146237],accel_mss,speed_ms,0,blend_radius_m)
  movel([0.578296, -1.177613, -2.695152, -0.839623, 1.570796, 2.149092],accel_mss,speed_ms,0,blend_radius_m)
  movel([0.580538, -1.179933, -2.694110, -0.838346, 1.570796, 2.151334],accel_mss,speed_ms,0,blend_radius_m)
  movel([0.582123, -1.182719, -2.692851, -0.836820, 1.570796, 2.152919],accel_mss,speed_ms,0,blend_radius_m)
  movel([0.583033, -1.185891, -2.691406, -0.835092, 1.570796, 2.153829],accel_mss,speed_ms,0,blend_radius_m)
  movel([0.583278, -1.189373, -2.689809, -0.833207, 1.570796, 2.154074],accel_mss,speed_ms,0,blend_radius_m)
  movel([0.582871, -1.193117, -2.688076, -0.831196, 1.570796, 2.153668],accel_mss,speed_ms,0,blend_radius_m)
  movel([0.581825, -1.197080, -2.686226, -0.829083, 1.570796, 2.152621],accel_mss,speed_ms,0,blend_radius_m)
  movel([0.580140, -1.201252, -2.684259, -0.826878, 1.570796, 2.150936],accel_mss,speed_ms,0,blend_radius_m)
  movel([0.579723, -1.202116, -2.683850, -0.826424, 1.570796, 2.150519],accel_mss,speed_ms,0,blend_radius_m)
  movel([0.581273, -1.202962, -2.683447, -0.825979, 1.570796, 2.152069],accel_mss,speed_ms,0,blend_radius_m)
  movel([0.583451, -1.204797, -2.682573, -0.825019, 1.570796, 2.154247],accel_mss,speed_ms,0,blend_radius_m)
  movel([0.584940, -1.206994, -2.681521, -0.823874, 1.570796, 2.155737],accel_mss,speed_ms,0,blend_radius_m)
  movel([0.585778, -1.209508, -2.680311, -0.822570, 1.570796, 2.156575],accel_mss,speed_ms,0,blend_radius_m)
  movel([0.585993, -1.212300, -2.678958, -0.821131, 1.570796, 2.156790],accel_mss,speed_ms,0,blend_radius_m)
  movel([0.585605, -1.215325, -2.677483, -0.819581, 1.570796, 2.156401],accel_mss,speed_ms,0,blend_radius_m)
  movel([0.584628, -1.218530, -2.675909, -0.817951, 1.570796, 2.155424],accel_mss,speed_ms,0,blend_radius_m)
  movel([0.583080, -1.221840, -2.674270, -0.816279, 1.570796, 2.153876],accel_mss,speed_ms,0,blend_radius_m)
  movel([0.580996, -1.225167, -2.672611, -0.814611, 1.570796, 2.151792],accel_mss,speed_ms,0,blend_radius_m)
  movel([0.578440, -1.228389, -2.670992, -0.813008, 1.570796, 2.149236],accel_mss,speed_ms,0,blend_radius_m)
  movel([0.575493, -1.231390, -2.669473, -0.811526, 1.570796, 2.146289],accel_mss,speed_ms,0,blend_radius_m)
  movel([0.572263, -1.234059, -2.668114, -0.810217, 1.570796, 2.143060],accel_mss,speed_ms,0,blend_radius_m)
  movel([0.568847, -1.236309, -2.666961, -0.809119, 1.570796, 2.139643],accel_mss,speed_ms,0,blend_radius_m)
  movel([0.565330, -1.238088, -2.666045, -0.808256, 1.570796, 2.136127],accel_mss,speed_ms,0,blend_radius_m)
  movel([0.561774, -1.239364, -2.665386, -0.807639, 1.570796, 2.132570],accel_mss,speed_ms,0,blend_radius_m)
  movel([0.558221, -1.240113, -2.664999, -0.807277, 1.570796, 2.129017],accel_mss,speed_ms,0,blend_radius_m)
  movel([0.554693, -1.240312, -2.664895, -0.807181, 1.570796, 2.125490],accel_mss,speed_ms,0,blend_radius_m)
  movel([0.554207, -1.240296, -2.664904, -0.807189, 1.570796, 2.125003],accel_mss,speed_ms,0,blend_radius_m)
  movel([0.552465, -1.241504, -2.664277, -0.806608, 1.570796, 2.123262],accel_mss,speed_ms,0,blend_radius_m)
  movel([0.549285, -1.244228, -2.662856, -0.805304, 1.570796, 2.120081],accel_mss,speed_ms,0,blend_radius_m)
  movel([0.547384, -1.245849, -2.662007, -0.804533, 1.570796, 2.118180],accel_mss,speed_ms,0,blend_radius_m)
  movel([0.545783, -1.247049, -2.661377, -0.803963, 1.570796, 2.116579],accel_mss,speed_ms,0,blend_radius_m)
  movel([0.542785, -1.248834, -2.660435, -0.803120, 1.570796, 2.113582],accel_mss,speed_ms,0,blend_radius_m)
  movel([0.539482, -1.250363, -2.659626, -0.802400, 1.570796, 2.110278],accel_mss,speed_ms,0,blend_radius_m)
  movel([0.536552, -1.251235, -2.659163, -0.801991, 1.570796, 2.107348],accel_mss,speed_ms,0,blend_radius_m)
  movel([0.533892, -1.251537, -2.659002, -0.801850, 1.570796, 2.104688],accel_mss,speed_ms,0,blend_radius_m)
  movel([0.531408, -1.251294, -2.659132, -0.801964, 1.570796, 2.102204],accel_mss,speed_ms,0,blend_radius_m)
  movel([0.529020, -1.250480, -2.659563, -0.802345, 1.570796, 2.099816],accel_mss,speed_ms,0,blend_radius_m)
  movel([0.526665, -1.249011, -2.660342, -0.803036, 1.570796, 2.097462],accel_mss,speed_ms,0,blend_radius_m)
  movel([0.524265, -1.246740, -2.661539, -0.804110, 1.570796, 2.095061],accel_mss,speed_ms,0,blend_radius_m)
  movel([0.521715, -1.243410, -2.663284, -0.805695, 1.570796, 2.092512],accel_mss,speed_ms,0,blend_radius_m)
  movel([0.518762, -1.238522, -2.665822, -0.808046, 1.570796, 2.089559],accel_mss,speed_ms,0,blend_radius_m)
  movel([0.514404, -1.230382, -2.669984, -0.812023, 1.570796, 2.085201],accel_mss,speed_ms,0,blend_radius_m)
  movel([0.510875, -1.224207, -2.673091, -0.815091, 1.570796, 2.081671],accel_mss,speed_ms,0,blend_radius_m)
  movel([0.508677, -1.220861, -2.674756, -0.816772, 1.570796, 2.079474],accel_mss,speed_ms,0,blend_radius_m)
  movel([0.506651, -1.218149, -2.676096, -0.818144, 1.570796, 2.077447],accel_mss,speed_ms,0,blend_radius_m)
  movel([0.504682, -1.215858, -2.677222, -0.819309, 1.570796, 2.075479],accel_mss,speed_ms,0,blend_radius_m)
  movel([0.502730, -1.213892, -2.678183, -0.820314, 1.570796, 2.073526],accel_mss,speed_ms,0,blend_radius_m)
  movel([0.500769, -1.212203, -2.679005, -0.821180, 1.570796, 2.071565],accel_mss,speed_ms,0,blend_radius_m)
  movel([0.498786, -1.210760, -2.679705, -0.821924, 1.570796, 2.069583],accel_mss,speed_ms,0,blend_radius_m)
  movel([0.494627, -1.208481, -2.680806, -0.823102, 1.570796, 2.065424],accel_mss,speed_ms,0,blend_radius_m)
  movel([0.490308, -1.207015, -2.681511, -0.823863, 1.570796, 2.061105],accel_mss,speed_ms,0,blend_radius_m)
  movel([0.485784, -1.206272, -2.681867, -0.824250, 1.570796, 2.056581],accel_mss,speed_ms,0,blend_radius_m)
  movel([0.481018, -1.206212, -2.681896, -0.824281, 1.570796, 2.051815],accel_mss,speed_ms,0,blend_radius_m)
  movel([0.479934, -1.206287, -2.681860, -0.824242, 1.570796, 2.050730],accel_mss,speed_ms,0,blend_radius_m)
  movel([0.477080, -1.206808, -2.681610, -0.823971, 1.570796, 2.047876],accel_mss,speed_ms,0,blend_radius_m)
  movel([0.472123, -1.208266, -2.680910, -0.823213, 1.570796, 2.042919],accel_mss,speed_ms,0,blend_radius_m)
  movel([0.469676, -1.209210, -2.680455, -0.822725, 1.570796, 2.040472],accel_mss,speed_ms,0,blend_radius_m)
  movel([0.467325, -1.210259, -2.679948, -0.822182, 1.570796, 2.038122],accel_mss,speed_ms,0,blend_radius_m)
  movel([0.465118, -1.211386, -2.679402, -0.821601, 1.570796, 2.035914],accel_mss,speed_ms,0,blend_radius_m)
  movel([0.463071, -1.212575, -2.678825, -0.820990, 1.570796, 2.033867],accel_mss,speed_ms,0,blend_radius_m)
  movel([0.461192, -1.213802, -2.678227, -0.820360, 1.570796, 2.031989],accel_mss,speed_ms,0,blend_radius_m)
  movel([0.459478, -1.215065, -2.677610, -0.819714, 1.570796, 2.030274],accel_mss,speed_ms,0,blend_radius_m)
  movel([0.457921, -1.216355, -2.676978, -0.819056, 1.570796, 2.028718],accel_mss,speed_ms,0,blend_radius_m)
  movel([0.455199, -1.219064, -2.675645, -0.817680, 1.570796, 2.025995],accel_mss,speed_ms,0,blend_radius_m)
  movel([0.453044, -1.221858, -2.674262, -0.816270, 1.570796, 2.023840],accel_mss,speed_ms,0,blend_radius_m)
  movel([0.452220, -1.223190, -2.673599, -0.815601, 1.570796, 2.023016],accel_mss,speed_ms,0,blend_radius_m)
  movel([0.451283, -1.225181, -2.672604, -0.814604, 1.570796, 2.022079],accel_mss,speed_ms,0,blend_radius_m)
  movel([0.450687, -1.227428, -2.671476, -0.813485, 1.570796, 2.021483],accel_mss,speed_ms,0,blend_radius_m)
  movel([0.450698, -1.229420, -2.670471, -0.812497, 1.570796, 2.021494],accel_mss,speed_ms,0,blend_radius_m)
  movel([0.451306, -1.231229, -2.669555, -0.811605, 1.570796, 2.022102],accel_mss,speed_ms,0,blend_radius_m)
  movel([0.452581, -1.232895, -2.668707, -0.810787, 1.570796, 2.023378],accel_mss,speed_ms,0,blend_radius_m)
  movel([0.454651, -1.234435, -2.667921, -0.810033, 1.570796, 2.025447],accel_mss,speed_ms,0,blend_radius_m)
  movel([0.457697, -1.235839, -2.667202, -0.809348, 1.570796, 2.028494],accel_mss,speed_ms,0,blend_radius_m)
  movel([0.461953, -1.237086, -2.666561, -0.808741, 1.570796, 2.032749],accel_mss,speed_ms,0,blend_radius_m)
  movel([0.467723, -1.238170, -2.666003, -0.808216, 1.570796, 2.038519],accel_mss,speed_ms,0,blend_radius_m)
  movel([0.475484, -1.239105, -2.665520, -0.807764, 1.570796, 2.046280],accel_mss,speed_ms,0,blend_radius_m)
  movel([0.486338, -1.240032, -2.665040, -0.807316, 1.570796, 2.057134],accel_mss,speed_ms,0,blend_radius_m)
  movel([0.494088, -1.240717, -2.664685, -0.806986, 1.570796, 2.064884],accel_mss,speed_ms,0,blend_radius_m)
  movel([0.500357, -1.241478, -2.664290, -0.806621, 1.570796, 2.071154],accel_mss,speed_ms,0,blend_radius_m)
  movel([0.503975, -1.242109, -2.663962, -0.806318, 1.570796, 2.074771],accel_mss,speed_ms,0,blend_radius_m)
  movel([0.506542, -1.242734, -2.663636, -0.806018, 1.570796, 2.077338],accel_mss,speed_ms,0,blend_radius_m)
  movel([0.508408, -1.243360, -2.663310, -0.805719, 1.570796, 2.079205],accel_mss,speed_ms,0,blend_radius_m)
  movel([0.510394, -1.244390, -2.662772, -0.805227, 1.570796, 2.081190],accel_mss,speed_ms,0,blend_radius_m)
  movel([0.511967, -1.245228, -2.662333, -0.804828, 1.570796, 2.082764],accel_mss,speed_ms,0,blend_radius_m)
  movel([0.513771, -1.246841, -2.661486, -0.804062, 1.570796, 2.084568],accel_mss,speed_ms,0,blend_radius_m)
  movel([0.515114, -1.248966, -2.660365, -0.803058, 1.570796, 2.085910],accel_mss,speed_ms,0,blend_radius_m)
  movel([0.515974, -1.251603, -2.658967, -0.801819, 1.570796, 2.086771],accel_mss,speed_ms,0,blend_radius_m)
  movel([0.516317, -1.254744, -2.657291, -0.800354, 1.570796, 2.087113],accel_mss,speed_ms,0,blend_radius_m)
  movel([0.516107, -1.258349, -2.655352, -0.798688, 1.570796, 2.086903],accel_mss,speed_ms,0,blend_radius_m)
  movel([0.515320, -1.262333, -2.653192, -0.796865, 1.570796, 2.086117],accel_mss,speed_ms,0,blend_radius_m)
  movel([0.513962, -1.266537, -2.650890, -0.794962, 1.570796, 2.084759],accel_mss,speed_ms,0,blend_radius_m)
  movel([0.512093, -1.270750, -2.648562, -0.793077, 1.570796, 2.082889],accel_mss,speed_ms,0,blend_radius_m)
  movel([0.510477, -1.273675, -2.646932, -0.791781, 1.570796, 2.081273],accel_mss,speed_ms,0,blend_radius_m)
  movel([0.508781, -1.276322, -2.645449, -0.790618, 1.570796, 2.079577],accel_mss,speed_ms,0,blend_radius_m)
  movel([0.506275, -1.279610, -2.643594, -0.789185, 1.570796, 2.077071],accel_mss,speed_ms,0,blend_radius_m)
  movel([0.503879, -1.282095, -2.642182, -0.788111, 1.570796, 2.074675],accel_mss,speed_ms,0,blend_radius_m)
  movel([0.501492, -1.284011, -2.641089, -0.787289, 1.570796, 2.072288],accel_mss,speed_ms,0,blend_radius_m)
  movel([0.498977, -1.285526, -2.640221, -0.786642, 1.570796, 2.069774],accel_mss,speed_ms,0,blend_radius_m)
  movel([0.496143, -1.286768, -2.639508, -0.786113, 1.570796, 2.066940],accel_mss,speed_ms,0,blend_radius_m)
  movel([0.492647, -1.287857, -2.638880, -0.785652, 1.570796, 2.063443],accel_mss,speed_ms,0,blend_radius_m)
  movel([0.487501, -1.289074, -2.638178, -0.785138, 1.570796, 2.058297],accel_mss,speed_ms,0,blend_radius_m)
  movel([0.480302, -1.290887, -2.637127, -0.784375, 1.570796, 2.051098],accel_mss,speed_ms,0,blend_radius_m)
  movel([0.479835, -1.291042, -2.637037, -0.784310, 1.570796, 2.050632],accel_mss,speed_ms,0,blend_radius_m)
  movel([0.480024, -1.291138, -2.636981, -0.784270, 1.570796, 2.050820],accel_mss,speed_ms,0,blend_radius_m)
  movel([0.482170, -1.291147, -2.636976, -0.784266, 1.570796, 2.052967],accel_mss,speed_ms,0,blend_radius_m)
  movel([0.490702, -1.290743, -2.637210, -0.784435, 1.570796, 2.061499],accel_mss,speed_ms,0,blend_radius_m)
  movel([0.501584, -1.290346, -2.637441, -0.784602, 1.570796, 2.072381],accel_mss,speed_ms,0,blend_radius_m)
  speed_ms = 0.05
  movel([0.501584, -1.234548, -2.609060, -0.868781, 1.570796, 2.072381],accel_mss,speed_ms,0,blend_radius_m)
  speed_ms = 0.051
  movel([0.501584, -1.224318, -2.603129, -0.884943, 1.570796, 2.072381],accel_mss,speed_ms,0,blend_radius_m)
  movel([0.490689, -1.263422, -2.581549, -0.867418, 1.570796, 2.061485],accel_mss,speed_ms,0,blend_radius_m)
  movel([0.490689, -1.294491, -2.598466, -0.819432, 1.570796, 2.061485],accel_mss,speed_ms,0,blend_radius_m)
  speed_ms = 0.017
  movel([0.490689, -1.328137, -2.614591, -0.769661, 1.570796, 2.061485],accel_mss,speed_ms,0,blend_radius_m)
  speed_ms = 0.051
  movel([0.489708, -1.330752, -2.612940, -0.768698, 1.570796, 2.060504],accel_mss,speed_ms,0,blend_radius_m)
  movel([0.489253, -1.333300, -2.611321, -0.767768, 1.570796, 2.060050],accel_mss,speed_ms,0,blend_radius_m)
  movel([0.489333, -1.335776, -2.609741, -0.766872, 1.570796, 2.060130],accel_mss,speed_ms,0,blend_radius_m)
  movel([0.489851, -1.337857, -2.608405, -0.766127, 1.570796, 2.060647],accel_mss,speed_ms,0,blend_radius_m)
  movel([0.492563, -1.334797, -2.610367, -0.767226, 1.570796, 2.063359],accel_mss,speed_ms,0,blend_radius_m)
  movel([0.495876, -1.331614, -2.612393, -0.768382, 1.570796, 2.066673],accel_mss,speed_ms,0,blend_radius_m)
  movel([0.499397, -1.328770, -2.614192, -0.769427, 1.570796, 2.070194],accel_mss,speed_ms,0,blend_radius_m)
  movel([0.503088, -1.326289, -2.615753, -0.770348, 1.570796, 2.073884],accel_mss,speed_ms,0,blend_radius_m)
  movel([0.506902, -1.324204, -2.617058, -0.771128, 1.570796, 2.077698],accel_mss,speed_ms,0,blend_radius_m)
  movel([0.510780, -1.322547, -2.618091, -0.771752, 1.570796, 2.081576],accel_mss,speed_ms,0,blend_radius_m)
  movel([0.514660, -1.321353, -2.618832, -0.772204, 1.570796, 2.085456],accel_mss,speed_ms,0,blend_radius_m)
  movel([0.518477, -1.320647, -2.619270, -0.772472, 1.570796, 2.089273],accel_mss,speed_ms,0,blend_radius_m)
  movel([0.522159, -1.320450, -2.619392, -0.772547, 1.570796, 2.092955],accel_mss,speed_ms,0,blend_radius_m)
  movel([0.525640, -1.320777, -2.619189, -0.772422, 1.570796, 2.096436],accel_mss,speed_ms,0,blend_radius_m)
  movel([0.528860, -1.321626, -2.618663, -0.772100, 1.570796, 2.099656],accel_mss,speed_ms,0,blend_radius_m)
  movel([0.531762, -1.322998, -2.617809, -0.771581, 1.570796, 2.102559],accel_mss,speed_ms,0,blend_radius_m)
  movel([0.534306, -1.324881, -2.616634, -0.770874, 1.570796, 2.105102],accel_mss,speed_ms,0,blend_radius_m)
  movel([0.535886, -1.326543, -2.615593, -0.770253, 1.570796, 2.106682],accel_mss,speed_ms,0,blend_radius_m)
  movel([0.537320, -1.329851, -2.613509, -0.769028, 1.570796, 2.108117],accel_mss,speed_ms,0,blend_radius_m)
  movel([0.538352, -1.333634, -2.611108, -0.767646, 1.570796, 2.109148],accel_mss,speed_ms,0,blend_radius_m)
  movel([0.538804, -1.337435, -2.608677, -0.766278, 1.570796, 2.109601],accel_mss,speed_ms,0,blend_radius_m)
  movel([0.538713, -1.341227, -2.606230, -0.764931, 1.570796, 2.109509],accel_mss,speed_ms,0,blend_radius_m)
  movel([0.538119, -1.344977, -2.603792, -0.763620, 1.570796, 2.108915],accel_mss,speed_ms,0,blend_radius_m)
  movel([0.537049, -1.348661, -2.601378, -0.762350, 1.570796, 2.107845],accel_mss,speed_ms,0,blend_radius_m)
  movel([0.535544, -1.352242, -2.599013, -0.761134, 1.570796, 2.106341],accel_mss,speed_ms,0,blend_radius_m)
  movel([0.533635, -1.355686, -2.596721, -0.759982, 1.570796, 2.104431],accel_mss,speed_ms,0,blend_radius_m)
  movel([0.531359, -1.358956, -2.594530, -0.758903, 1.570796, 2.102156],accel_mss,speed_ms,0,blend_radius_m)
  movel([0.528758, -1.362012, -2.592469, -0.757909, 1.570796, 2.099554],accel_mss,speed_ms,0,blend_radius_m)
  movel([0.525880, -1.364812, -2.590569, -0.757009, 1.570796, 2.096677],accel_mss,speed_ms,0,blend_radius_m)
  movel([0.522773, -1.367314, -2.588861, -0.756214, 1.570796, 2.093569],accel_mss,speed_ms,0,blend_radius_m)
  movel([0.519494, -1.369480, -2.587375, -0.755533, 1.570796, 2.090291],accel_mss,speed_ms,0,blend_radius_m)
  movel([0.516097, -1.371282, -2.586135, -0.754972, 1.570796, 2.086893],accel_mss,speed_ms,0,blend_radius_m)
  movel([0.512626, -1.372693, -2.585160, -0.754536, 1.570796, 2.083422],accel_mss,speed_ms,0,blend_radius_m)
  movel([0.509133, -1.373690, -2.584469, -0.754230, 1.570796, 2.079929],accel_mss,speed_ms,0,blend_radius_m)
  movel([0.505647, -1.374263, -2.584072, -0.754054, 1.570796, 2.076444],accel_mss,speed_ms,0,blend_radius_m)
  movel([0.502209, -1.374392, -2.583982, -0.754015, 1.570796, 2.073006],accel_mss,speed_ms,0,blend_radius_m)
  movel([0.498837, -1.374065, -2.584209, -0.754115, 1.570796, 2.069634],accel_mss,speed_ms,0,blend_radius_m)
  movel([0.495560, -1.373257, -2.584769, -0.754363, 1.570796, 2.066356],accel_mss,speed_ms,0,blend_radius_m)
  movel([0.492398, -1.371950, -2.585674, -0.754766, 1.570796, 2.063195],accel_mss,speed_ms,0,blend_radius_m)
  movel([0.489377, -1.370111, -2.586942, -0.755337, 1.570796, 2.060174],accel_mss,speed_ms,0,blend_radius_m)
  movel([0.486524, -1.367710, -2.588590, -0.756089, 1.570796, 2.057320],accel_mss,speed_ms,0,blend_radius_m)
  movel([0.483859, -1.364710, -2.590638, -0.757041, 1.570796, 2.054655],accel_mss,speed_ms,0,blend_radius_m)
  movel([0.481419, -1.361062, -2.593111, -0.758216, 1.570796, 2.052215],accel_mss,speed_ms,0,blend_radius_m)
  movel([0.479236, -1.356722, -2.596029, -0.759639, 1.570796, 2.050032],accel_mss,speed_ms,0,blend_radius_m)
  movel([0.477345, -1.351637, -2.599414, -0.761339, 1.570796, 2.048141],accel_mss,speed_ms,0,blend_radius_m)
  movel([0.476142, -1.347286, -2.602281, -0.762822, 1.570796, 2.046938],accel_mss,speed_ms,0,blend_radius_m)
  movel([0.475310, -1.343058, -2.605043, -0.764289, 1.570796, 2.046106],accel_mss,speed_ms,0,blend_radius_m)
  movel([0.474768, -1.337816, -2.608432, -0.766141, 1.570796, 2.045564],accel_mss,speed_ms,0,blend_radius_m)
  movel([0.474790, -1.332897, -2.611578, -0.767914, 1.570796, 2.045586],accel_mss,speed_ms,0,blend_radius_m)
  movel([0.475330, -1.328281, -2.614500, -0.769608, 1.570796, 2.046126],accel_mss,speed_ms,0,blend_radius_m)
  movel([0.476334, -1.323950, -2.617216, -0.771223, 1.570796, 2.047130],accel_mss,speed_ms,0,blend_radius_m)
  movel([0.477770, -1.319875, -2.619748, -0.772766, 1.570796, 2.048566],accel_mss,speed_ms,0,blend_radius_m)
  movel([0.479600, -1.316044, -2.622109, -0.774237, 1.570796, 2.050396],accel_mss,speed_ms,0,blend_radius_m)
  movel([0.481811, -1.312430, -2.624317, -0.775642, 1.570796, 2.052607],accel_mss,speed_ms,0,blend_radius_m)
  movel([0.484390, -1.309014, -2.626389, -0.776986, 1.570796, 2.055186],accel_mss,speed_ms,0,blend_radius_m)
  movel([0.487335, -1.305787, -2.628332, -0.778270, 1.570796, 2.058131],accel_mss,speed_ms,0,blend_radius_m)
  movel([0.490659, -1.302739, -2.630154, -0.779496, 1.570796, 2.061456],accel_mss,speed_ms,0,blend_radius_m)
  movel([0.494366, -1.299885, -2.631850, -0.780654, 1.570796, 2.065162],accel_mss,speed_ms,0,blend_radius_m)
  movel([0.498457, -1.297240, -2.633412, -0.781737, 1.570796, 2.069253],accel_mss,speed_ms,0,blend_radius_m)
  movel([0.502924, -1.294843, -2.634820, -0.782726, 1.570796, 2.073721],accel_mss,speed_ms,0,blend_radius_m)
  movel([0.507728, -1.292743, -2.636047, -0.783599, 1.570796, 2.078525],accel_mss,speed_ms,0,blend_radius_m)
  movel([0.512790, -1.291013, -2.637054, -0.784322, 1.570796, 2.083586],accel_mss,speed_ms,0,blend_radius_m)
  movel([0.517984, -1.289721, -2.637803, -0.784865, 1.570796, 2.088780],accel_mss,speed_ms,0,blend_radius_m)
  movel([0.523127, -1.288939, -2.638255, -0.785194, 1.570796, 2.093923],accel_mss,speed_ms,0,blend_radius_m)
  movel([0.527990, -1.288708, -2.638389, -0.785292, 1.570796, 2.098786],accel_mss,speed_ms,0,blend_radius_m)
  movel([0.532330, -1.289034, -2.638201, -0.785155, 1.570796, 2.103126],accel_mss,speed_ms,0,blend_radius_m)
  movel([0.535949, -1.289864, -2.637720, -0.784805, 1.570796, 2.106745],accel_mss,speed_ms,0,blend_radius_m)
  movel([0.538594, -1.291024, -2.637047, -0.784318, 1.570796, 2.109390],accel_mss,speed_ms,0,blend_radius_m)
  movel([0.541413, -1.291862, -2.636560, -0.783967, 1.570796, 2.112209],accel_mss,speed_ms,0,blend_radius_m)
  movel([0.546703, -1.293936, -2.635350, -0.783103, 1.570796, 2.117499],accel_mss,speed_ms,0,blend_radius_m)
  movel([0.554400, -1.297544, -2.633233, -0.781612, 1.570796, 2.125196],accel_mss,speed_ms,0,blend_radius_m)
  movel([0.561304, -1.300717, -2.631357, -0.780315, 1.570796, 2.132100],accel_mss,speed_ms,0,blend_radius_m)
  movel([0.564166, -1.301831, -2.630695, -0.779863, 1.570796, 2.134963],accel_mss,speed_ms,0,blend_radius_m)
  movel([0.566479, -1.302572, -2.630254, -0.779563, 1.570796, 2.137275],accel_mss,speed_ms,0,blend_radius_m)
  movel([0.568442, -1.303049, -2.629969, -0.779371, 1.570796, 2.139239],accel_mss,speed_ms,0,blend_radius_m)
  movel([0.570146, -1.303316, -2.629810, -0.779263, 1.570796, 2.140942],accel_mss,speed_ms,0,blend_radius_m)
  movel([0.571644, -1.303415, -2.629751, -0.779223, 1.570796, 2.142440],accel_mss,speed_ms,0,blend_radius_m)
  movel([0.572973, -1.303368, -2.629779, -0.779242, 1.570796, 2.143769],accel_mss,speed_ms,0,blend_radius_m)
  movel([0.574167, -1.303199, -2.629880, -0.779310, 1.570796, 2.144963],accel_mss,speed_ms,0,blend_radius_m)
  movel([0.575243, -1.302925, -2.630043, -0.779421, 1.570796, 2.146039],accel_mss,speed_ms,0,blend_radius_m)
  movel([0.577176, -1.302074, -2.630550, -0.779764, 1.570796, 2.147973],accel_mss,speed_ms,0,blend_radius_m)
  movel([0.578841, -1.300864, -2.631269, -0.780255, 1.570796, 2.149637],accel_mss,speed_ms,0,blend_radius_m)
  movel([0.580080, -1.299577, -2.632032, -0.780780, 1.570796, 2.150876],accel_mss,speed_ms,0,blend_radius_m)
  movel([0.581511, -1.297397, -2.633320, -0.781673, 1.570796, 2.152307],accel_mss,speed_ms,0,blend_radius_m)
  movel([0.582449, -1.295239, -2.634588, -0.782562, 1.570796, 2.153245],accel_mss,speed_ms,0,blend_radius_m)
  movel([0.582913, -1.293050, -2.635868, -0.783471, 1.570796, 2.153709],accel_mss,speed_ms,0,blend_radius_m)
  movel([0.582918, -1.290657, -2.637260, -0.784472, 1.570796, 2.153714],accel_mss,speed_ms,0,blend_radius_m)
  movel([0.582396, -1.287762, -2.638935, -0.785692, 1.570796, 2.153193],accel_mss,speed_ms,0,blend_radius_m)
  movel([0.581111, -1.283421, -2.641426, -0.787542, 1.570796, 2.151908],accel_mss,speed_ms,0,blend_radius_m)
  movel([0.579823, -1.278570, -2.644182, -0.789637, 1.570796, 2.150620],accel_mss,speed_ms,0,blend_radius_m)
  movel([0.579433, -1.276230, -2.645501, -0.790658, 1.570796, 2.150229],accel_mss,speed_ms,0,blend_radius_m)
  movel([0.579237, -1.274051, -2.646722, -0.791615, 1.570796, 2.150034],accel_mss,speed_ms,0,blend_radius_m)
  movel([0.579207, -1.271928, -2.647907, -0.792554, 1.570796, 2.150003],accel_mss,speed_ms,0,blend_radius_m)
  movel([0.579326, -1.269815, -2.649080, -0.793493, 1.570796, 2.150123],accel_mss,speed_ms,0,blend_radius_m)
  movel([0.580039, -1.265414, -2.651507, -0.795468, 1.570796, 2.150835],accel_mss,speed_ms,0,blend_radius_m)
  movel([0.581375, -1.260818, -2.654015, -0.797555, 1.570796, 2.152171],accel_mss,speed_ms,0,blend_radius_m)
  movel([0.582506, -1.257883, -2.655604, -0.798902, 1.570796, 2.153302],accel_mss,speed_ms,0,blend_radius_m)
  movel([0.587495, -1.249354, -2.660160, -0.802875, 1.570796, 2.158291],accel_mss,speed_ms,0,blend_radius_m)
  movel([0.588735, -1.247049, -2.661377, -0.803963, 1.570796, 2.159532],accel_mss,speed_ms,0,blend_radius_m)
  movel([0.589174, -1.245966, -2.661946, -0.804477, 1.570796, 2.159971],accel_mss,speed_ms,0,blend_radius_m)
  movel([0.589485, -1.244213, -2.662864, -0.805311, 1.570796, 2.160281],accel_mss,speed_ms,0,blend_radius_m)
  movel([0.589364, -1.241475, -2.664292, -0.806622, 1.570796, 2.160160],accel_mss,speed_ms,0,blend_radius_m)
  movel([0.589119, -1.234223, -2.668030, -0.810136, 1.570796, 2.159916],accel_mss,speed_ms,0,blend_radius_m)
  movel([0.589709, -1.232124, -2.669100, -0.811165, 1.570796, 2.160505],accel_mss,speed_ms,0,blend_radius_m)
  movel([0.590927, -1.229554, -2.670404, -0.812432, 1.570796, 2.161723],accel_mss,speed_ms,0,blend_radius_m)
  movel([0.593038, -1.225991, -2.672198, -0.814200, 1.570796, 2.163835],accel_mss,speed_ms,0,blend_radius_m)
  movel([0.594405, -1.223696, -2.673346, -0.815347, 1.570796, 2.165201],accel_mss,speed_ms,0,blend_radius_m)
  movel([0.595399, -1.221795, -2.674293, -0.816301, 1.570796, 2.166195],accel_mss,speed_ms,0,blend_radius_m)
  movel([0.595975, -1.220411, -2.674979, -0.816999, 1.570796, 2.166771],accel_mss,speed_ms,0,blend_radius_m)
  movel([0.596313, -1.219243, -2.675557, -0.817589, 1.570796, 2.167110],accel_mss,speed_ms,0,blend_radius_m)
  movel([0.596459, -1.217266, -2.676531, -0.818592, 1.570796, 2.167255],accel_mss,speed_ms,0,blend_radius_m)
  movel([0.596887, -1.218693, -2.675828, -0.817868, 1.570796, 2.167683],accel_mss,speed_ms,0,blend_radius_m)
  movel([0.596951, -1.220853, -2.674760, -0.816776, 1.570796, 2.167748],accel_mss,speed_ms,0,blend_radius_m)
  movel([0.596454, -1.223374, -2.673507, -0.815508, 1.570796, 2.167251],accel_mss,speed_ms,0,blend_radius_m)
  movel([0.595331, -1.226518, -2.671933, -0.813937, 1.570796, 2.166128],accel_mss,speed_ms,0,blend_radius_m)
  movel([0.593271, -1.231228, -2.669555, -0.811606, 1.570796, 2.164067],accel_mss,speed_ms,0,blend_radius_m)
  movel([0.592118, -1.234143, -2.668070, -0.810175, 1.570796, 2.162914],accel_mss,speed_ms,0,blend_radius_m)
  movel([0.591591, -1.235881, -2.667181, -0.809328, 1.570796, 2.162387],accel_mss,speed_ms,0,blend_radius_m)
  movel([0.591303, -1.237310, -2.666446, -0.808633, 1.570796, 2.162099],accel_mss,speed_ms,0,blend_radius_m)
  movel([0.591199, -1.238558, -2.665803, -0.808028, 1.570796, 2.161995],accel_mss,speed_ms,0,blend_radius_m)
  movel([0.591483, -1.240757, -2.664665, -0.806967, 1.570796, 2.162280],accel_mss,speed_ms,0,blend_radius_m)
  movel([0.592411, -1.242611, -2.663701, -0.806077, 1.570796, 2.163208],accel_mss,speed_ms,0,blend_radius_m)
  movel([0.592513, -1.242748, -2.663629, -0.806012, 1.570796, 2.163309],accel_mss,speed_ms,0,blend_radius_m)
  movel([0.595525, -1.241871, -2.664086, -0.806432, 1.570796, 2.166322],accel_mss,speed_ms,0,blend_radius_m)
  movel([0.597693, -1.241703, -2.664173, -0.806513, 1.570796, 2.168490],accel_mss,speed_ms,0,blend_radius_m)
  movel([0.599125, -1.242109, -2.663962, -0.806318, 1.570796, 2.169921],accel_mss,speed_ms,0,blend_radius_m)
  movel([0.600072, -1.243013, -2.663491, -0.805885, 1.570796, 2.170868],accel_mss,speed_ms,0,blend_radius_m)
  movel([0.600669, -1.244511, -2.662709, -0.805169, 1.570796, 2.171466],accel_mss,speed_ms,0,blend_radius_m)
  movel([0.601008, -1.246995, -2.661405, -0.803989, 1.570796, 2.171804],accel_mss,speed_ms,0,blend_radius_m)
  movel([0.601277, -1.250011, -2.659812, -0.802566, 1.570796, 2.172073],accel_mss,speed_ms,0,blend_radius_m)
  movel([0.602500, -1.253646, -2.657879, -0.800865, 1.570796, 2.173296],accel_mss,speed_ms,0,blend_radius_m)
  movel([0.604855, -1.260075, -2.654419, -0.797895, 1.570796, 2.175652],accel_mss,speed_ms,0,blend_radius_m)
  movel([0.605314, -1.262059, -2.653341, -0.796990, 1.570796, 2.176110],accel_mss,speed_ms,0,blend_radius_m)
  movel([0.605598, -1.264738, -2.651878, -0.795774, 1.570796, 2.176394],accel_mss,speed_ms,0,blend_radius_m)
  movel([0.605504, -1.267071, -2.650596, -0.794722, 1.570796, 2.176301],accel_mss,speed_ms,0,blend_radius_m)
  movel([0.604900, -1.270526, -2.648686, -0.793177, 1.570796, 2.175696],accel_mss,speed_ms,0,blend_radius_m)
  movel([0.603669, -1.274915, -2.646239, -0.791235, 1.570796, 2.174466],accel_mss,speed_ms,0,blend_radius_m)
  movel([0.601404, -1.282148, -2.642153, -0.788089, 1.570796, 2.172200],accel_mss,speed_ms,0,blend_radius_m)
  movel([0.600919, -1.284115, -2.641030, -0.787244, 1.570796, 2.171715],accel_mss,speed_ms,0,blend_radius_m)
  movel([0.600192, -1.288118, -2.638729, -0.785541, 1.570796, 2.170988],accel_mss,speed_ms,0,blend_radius_m)
  movel([0.599470, -1.293752, -2.635458, -0.783179, 1.570796, 2.170266],accel_mss,speed_ms,0,blend_radius_m)
  movel([0.598967, -1.296770, -2.633688, -0.781930, 1.570796, 2.169764],accel_mss,speed_ms,0,blend_radius_m)
  movel([0.598494, -1.298665, -2.632571, -0.781152, 1.570796, 2.169290],accel_mss,speed_ms,0,blend_radius_m)
  movel([0.597940, -1.300333, -2.631584, -0.780471, 1.570796, 2.168737],accel_mss,speed_ms,0,blend_radius_m)
  movel([0.597282, -1.301922, -2.630641, -0.779826, 1.570796, 2.168079],accel_mss,speed_ms,0,blend_radius_m)
  movel([0.595532, -1.305165, -2.628705, -0.778519, 1.570796, 2.166329],accel_mss,speed_ms,0,blend_radius_m)
  movel([0.593095, -1.308680, -2.626590, -0.777118, 1.570796, 2.163891],accel_mss,speed_ms,0,blend_radius_m)
  movel([0.590150, -1.312267, -2.624416, -0.775706, 1.570796, 2.160947],accel_mss,speed_ms,0,blend_radius_m)
  movel([0.586214, -1.316458, -2.621854, -0.774077, 1.570796, 2.157011],accel_mss,speed_ms,0,blend_radius_m)
  movel([0.582582, -1.319774, -2.619811, -0.772805, 1.570796, 2.153379],accel_mss,speed_ms,0,blend_radius_m)
  movel([0.579139, -1.322407, -2.618178, -0.771805, 1.570796, 2.149935],accel_mss,speed_ms,0,blend_radius_m)
  movel([0.575831, -1.324464, -2.616895, -0.771030, 1.570796, 2.146627],accel_mss,speed_ms,0,blend_radius_m)
  movel([0.572601, -1.326022, -2.615920, -0.770447, 1.570796, 2.143397],accel_mss,speed_ms,0,blend_radius_m)
  movel([0.569389, -1.327137, -2.615220, -0.770032, 1.570796, 2.140185],accel_mss,speed_ms,0,blend_radius_m)
  movel([0.566130, -1.327832, -2.614783, -0.769774, 1.570796, 2.136927],accel_mss,speed_ms,0,blend_radius_m)
  movel([0.562757, -1.328108, -2.614609, -0.769672, 1.570796, 2.133553],accel_mss,speed_ms,0,blend_radius_m)
  movel([0.559196, -1.327942, -2.614714, -0.769733, 1.570796, 2.129993],accel_mss,speed_ms,0,blend_radius_m)
  movel([0.555361, -1.327282, -2.615129, -0.769978, 1.570796, 2.126157],accel_mss,speed_ms,0,blend_radius_m)
  movel([0.551122, -1.326050, -2.615902, -0.770437, 1.570796, 2.121918],accel_mss,speed_ms,0,blend_radius_m)
  movel([0.546261, -1.324125, -2.617107, -0.771157, 1.570796, 2.117057],accel_mss,speed_ms,0,blend_radius_m)
  movel([0.540244, -1.321255, -2.618893, -0.772241, 1.570796, 2.111040],accel_mss,speed_ms,0,blend_radius_m)
  movel([0.530412, -1.316374, -2.621906, -0.774109, 1.570796, 2.101209],accel_mss,speed_ms,0,blend_radius_m)
  movel([0.526696, -1.314776, -2.622885, -0.774728, 1.570796, 2.097492],accel_mss,speed_ms,0,blend_radius_m)
  movel([0.523808, -1.313728, -2.623525, -0.775135, 1.570796, 2.094604],accel_mss,speed_ms,0,blend_radius_m)
  movel([0.521314, -1.312998, -2.623971, -0.775420, 1.570796, 2.092110],accel_mss,speed_ms,0,blend_radius_m)
  movel([0.519070, -1.312504, -2.624272, -0.775613, 1.570796, 2.089867],accel_mss,speed_ms,0,blend_radius_m)
  movel([0.517018, -1.312204, -2.624454, -0.775730, 1.570796, 2.087815],accel_mss,speed_ms,0,blend_radius_m)
  movel([0.515110, -1.312069, -2.624537, -0.775784, 1.570796, 2.085906],accel_mss,speed_ms,0,blend_radius_m)
  movel([0.513321, -1.312081, -2.624529, -0.775779, 1.570796, 2.084118],accel_mss,speed_ms,0,blend_radius_m)
  movel([0.511632, -1.312223, -2.624443, -0.775723, 1.570796, 2.082428],accel_mss,speed_ms,0,blend_radius_m)
  movel([0.508414, -1.312883, -2.624041, -0.775465, 1.570796, 2.079210],accel_mss,speed_ms,0,blend_radius_m)
  movel([0.505446, -1.313980, -2.623372, -0.775037, 1.570796, 2.076242],accel_mss,speed_ms,0,blend_radius_m)
  movel([0.502636, -1.315495, -2.622445, -0.774449, 1.570796, 2.073433],accel_mss,speed_ms,0,blend_radius_m)
  movel([0.499902, -1.317457, -2.621240, -0.773692, 1.570796, 2.070698],accel_mss,speed_ms,0,blend_radius_m)
  movel([0.497188, -1.319916, -2.619723, -0.772750, 1.570796, 2.067985],accel_mss,speed_ms,0,blend_radius_m)
  movel([0.494443, -1.322968, -2.617828, -0.771593, 1.570796, 2.065239],accel_mss,speed_ms,0,blend_radius_m)
  movel([0.491636, -1.326718, -2.615483, -0.770188, 1.570796, 2.062432],accel_mss,speed_ms,0,blend_radius_m)
  movel([0.490689, -1.328137, -2.614591, -0.769661, 1.570796, 2.061485],accel_mss,speed_ms,0,blend_radius_m)
  speed_ms = 0.05
  movel([0.490689, -1.273498, -2.587272, -0.851619, 1.570796, 2.061485],accel_mss,speed_ms,0,blend_radius_m)
  speed_ms = 0.051
  movel([0.490689, -1.263422, -2.581549, -0.867418, 1.570796, 2.061485],accel_mss,speed_ms,0,blend_radius_m)
  movel([0.589787, -1.201739, -2.614801, -0.895849, 1.570796, 2.160584],accel_mss,speed_ms,0,blend_radius_m)
  movel([0.589787, -1.233601, -2.632710, -0.846078, 1.570796, 2.160584],accel_mss,speed_ms,0,blend_radius_m)
  speed_ms = 0.017
  movel([0.589787, -1.268422, -2.649851, -0.794116, 1.570796, 2.160584],accel_mss,speed_ms,0,blend_radius_m)
  speed_ms = 0.051
  movel([0.590529, -1.268191, -2.649979, -0.794219, 1.570796, 2.161325],accel_mss,speed_ms,0,blend_radius_m)
  movel([0.590837, -1.268341, -2.649896, -0.794152, 1.570796, 2.161633],accel_mss,speed_ms,0,blend_radius_m)
  movel([0.590849, -1.268352, -2.649890, -0.794147, 1.570796, 2.161645],accel_mss,speed_ms,0,blend_radius_m)
  movel([0.591531, -1.268843, -2.649618, -0.793927, 1.570796, 2.162328],accel_mss,speed_ms,0,blend_radius_m)
  movel([0.592437, -1.268762, -2.649663, -0.793964, 1.570796, 2.163234],accel_mss,speed_ms,0,blend_radius_m)
  movel([0.593675, -1.268155, -2.649999, -0.794236, 1.570796, 2.164472],accel_mss,speed_ms,0,blend_radius_m)
  movel([0.595420, -1.266885, -2.650699, -0.794805, 1.570796, 2.166216],accel_mss,speed_ms,0,blend_radius_m)
  movel([0.596672, -1.265858, -2.651263, -0.795268, 1.570796, 2.167468],accel_mss,speed_ms,0,blend_radius_m)
  movel([0.596966, -1.265623, -2.651392, -0.795374, 1.570796, 2.167762],accel_mss,speed_ms,0,blend_radius_m)
  movel([0.596854, -1.264255, -2.652142, -0.795992, 1.570796, 2.167650],accel_mss,speed_ms,0,blend_radius_m)
  movel([0.596613, -1.263247, -2.652693, -0.796449, 1.570796, 2.167409],accel_mss,speed_ms,0,blend_radius_m)
  movel([0.596310, -1.262578, -2.653058, -0.796753, 1.570796, 2.167106],accel_mss,speed_ms,0,blend_radius_m)
  movel([0.595897, -1.262065, -2.653338, -0.796987, 1.570796, 2.166694],accel_mss,speed_ms,0,blend_radius_m)
  movel([0.595417, -1.261746, -2.653511, -0.797132, 1.570796, 2.166213],accel_mss,speed_ms,0,blend_radius_m)
  movel([0.594226, -1.261585, -2.653599, -0.797206, 1.570796, 2.165022],accel_mss,speed_ms,0,blend_radius_m)
  movel([0.592713, -1.262029, -2.653357, -0.797003, 1.570796, 2.163509],accel_mss,speed_ms,0,blend_radius_m)
  movel([0.591336, -1.262769, -2.652954, -0.796666, 1.570796, 2.162132],accel_mss,speed_ms,0,blend_radius_m)
  movel([0.592047, -1.260939, -2.653950, -0.797500, 1.570796, 2.162843],accel_mss,speed_ms,0,blend_radius_m)
  movel([0.592604, -1.259910, -2.654508, -0.797971, 1.570796, 2.163401],accel_mss,speed_ms,0,blend_radius_m)
  movel([0.592930, -1.259521, -2.654718, -0.798149, 1.570796, 2.163726],accel_mss,speed_ms,0,blend_radius_m)
  movel([0.593285, -1.259257, -2.654861, -0.798270, 1.570796, 2.164081],accel_mss,speed_ms,0,blend_radius_m)
  movel([0.594052, -1.259121, -2.654935, -0.798333, 1.570796, 2.164848],accel_mss,speed_ms,0,blend_radius_m)
  movel([0.594734, -1.259365, -2.654803, -0.798221, 1.570796, 2.165530],accel_mss,speed_ms,0,blend_radius_m)
  movel([0.596536, -1.260763, -2.654045, -0.797581, 1.570796, 2.167333],accel_mss,speed_ms,0,blend_radius_m)
  movel([0.597139, -1.261510, -2.653639, -0.797239, 1.570796, 2.167935],accel_mss,speed_ms,0,blend_radius_m)
  movel([0.597620, -1.262345, -2.653185, -0.796859, 1.570796, 2.168417],accel_mss,speed_ms,0,blend_radius_m)
  movel([0.597947, -1.263254, -2.652689, -0.796446, 1.570796, 2.168743],accel_mss,speed_ms,0,blend_radius_m)
  movel([0.598093, -1.264150, -2.652200, -0.796040, 1.570796, 2.168889],accel_mss,speed_ms,0,blend_radius_m)
  movel([0.598072, -1.265026, -2.651720, -0.795643, 1.570796, 2.168868],accel_mss,speed_ms,0,blend_radius_m)
  movel([0.597909, -1.265877, -2.651253, -0.795259, 1.570796, 2.168705],accel_mss,speed_ms,0,blend_radius_m)
  movel([0.597157, -1.267562, -2.650326, -0.794501, 1.570796, 2.167954],accel_mss,speed_ms,0,blend_radius_m)
  movel([0.596724, -1.268199, -2.649974, -0.794216, 1.570796, 2.167520],accel_mss,speed_ms,0,blend_radius_m)
  movel([0.595521, -1.267353, -2.650441, -0.794595, 1.570796, 2.166317],accel_mss,speed_ms,0,blend_radius_m)
  movel([0.593551, -1.273044, -2.647285, -0.792060, 1.570796, 2.164348],accel_mss,speed_ms,0,blend_radius_m)
  movel([0.593496, -1.273207, -2.647194, -0.791988, 1.570796, 2.164292],accel_mss,speed_ms,0,blend_radius_m)
  movel([0.592073, -1.272864, -2.647385, -0.792139, 1.570796, 2.162869],accel_mss,speed_ms,0,blend_radius_m)
  movel([0.591043, -1.272040, -2.647845, -0.792504, 1.570796, 2.161839],accel_mss,speed_ms,0,blend_radius_m)
  movel([0.590312, -1.270665, -2.648609, -0.793115, 1.570796, 2.161108],accel_mss,speed_ms,0,blend_radius_m)
  movel([0.589801, -1.268510, -2.649802, -0.794076, 1.570796, 2.160597],accel_mss,speed_ms,0,blend_radius_m)
  movel([0.589787, -1.268422, -2.649851, -0.794116, 1.570796, 2.160584],accel_mss,speed_ms,0,blend_radius_m)
  speed_ms = 0.05
  movel([0.589787, -1.212040, -2.620852, -0.879497, 1.570796, 2.160584],accel_mss,speed_ms,0,blend_radius_m)
  speed_ms = 0.051
  movel([0.589787, -1.201739, -2.614801, -0.895849, 1.570796, 2.160584],accel_mss,speed_ms,0,blend_radius_m)
  movel([0.521520, -1.275543, -2.574496, -0.862350, 1.570796, 2.092316],accel_mss,speed_ms,0,blend_radius_m)
  movel([0.521520, -1.306424, -2.591219, -0.814746, 1.570796, 2.092316],accel_mss,speed_ms,0,blend_radius_m)
  speed_ms = 0.017
  movel([0.521520, -1.339809, -2.607147, -0.765432, 1.570796, 2.092316],accel_mss,speed_ms,0,blend_radius_m)
  speed_ms = 0.051
  movel([0.520353, -1.338539, -2.607966, -0.765883, 1.570796, 2.091149],accel_mss,speed_ms,0,blend_radius_m)
  movel([0.518935, -1.337848, -2.608411, -0.766130, 1.570796, 2.089732],accel_mss,speed_ms,0,blend_radius_m)
  movel([0.517283, -1.337660, -2.608532, -0.766197, 1.570796, 2.088079],accel_mss,speed_ms,0,blend_radius_m)
  movel([0.515386, -1.337948, -2.608347, -0.766094, 1.570796, 2.086183],accel_mss,speed_ms,0,blend_radius_m)
  movel([0.513217, -1.338730, -2.607843, -0.765816, 1.570796, 2.084013],accel_mss,speed_ms,0,blend_radius_m)
  movel([0.510773, -1.340049, -2.606992, -0.765347, 1.570796, 2.081569],accel_mss,speed_ms,0,blend_radius_m)
  movel([0.508098, -1.341936, -2.605771, -0.764682, 1.570796, 2.078894],accel_mss,speed_ms,0,blend_radius_m)
  movel([0.505330, -1.344355, -2.604198, -0.763836, 1.570796, 2.076126],accel_mss,speed_ms,0,blend_radius_m)
  movel([0.502716, -1.347141, -2.602376, -0.762872, 1.570796, 2.073513],accel_mss,speed_ms,0,blend_radius_m)
  movel([0.500548, -1.350008, -2.600490, -0.761891, 1.570796, 2.071345],accel_mss,speed_ms,0,blend_radius_m)
  movel([0.499059, -1.352632, -2.598754, -0.761003, 1.570796, 2.069855],accel_mss,speed_ms,0,blend_radius_m)
  movel([0.498589, -1.353786, -2.597988, -0.760616, 1.570796, 2.069386],accel_mss,speed_ms,0,blend_radius_m)
  movel([0.500673, -1.354917, -2.597234, -0.760238, 1.570796, 2.071469],accel_mss,speed_ms,0,blend_radius_m)
  movel([0.502090, -1.355482, -2.596857, -0.760050, 1.570796, 2.072887],accel_mss,speed_ms,0,blend_radius_m)
  movel([0.503516, -1.355901, -2.596577, -0.759910, 1.570796, 2.074313],accel_mss,speed_ms,0,blend_radius_m)
  movel([0.504921, -1.356175, -2.596394, -0.759820, 1.570796, 2.075717],accel_mss,speed_ms,0,blend_radius_m)
  movel([0.506289, -1.356310, -2.596304, -0.759775, 1.570796, 2.077086],accel_mss,speed_ms,0,blend_radius_m)
  movel([0.507609, -1.356316, -2.596300, -0.759773, 1.570796, 2.078406],accel_mss,speed_ms,0,blend_radius_m)
  movel([0.508877, -1.356203, -2.596376, -0.759810, 1.570796, 2.079673],accel_mss,speed_ms,0,blend_radius_m)
  movel([0.511321, -1.355632, -2.596757, -0.760000, 1.570796, 2.082118],accel_mss,speed_ms,0,blend_radius_m)
  movel([0.513567, -1.354656, -2.597408, -0.760325, 1.570796, 2.084364],accel_mss,speed_ms,0,blend_radius_m)
  movel([0.515665, -1.353295, -2.598314, -0.760780, 1.570796, 2.086461],accel_mss,speed_ms,0,blend_radius_m)
  movel([0.517666, -1.351514, -2.599495, -0.761380, 1.570796, 2.088462],accel_mss,speed_ms,0,blend_radius_m)
  movel([0.519120, -1.349869, -2.600582, -0.761938, 1.570796, 2.089917],accel_mss,speed_ms,0,blend_radius_m)
  movel([0.520131, -1.348503, -2.601481, -0.762404, 1.570796, 2.090928],accel_mss,speed_ms,0,blend_radius_m)
  movel([0.521439, -1.346212, -2.602985, -0.763192, 1.570796, 2.092235],accel_mss,speed_ms,0,blend_radius_m)
  movel([0.522155, -1.344110, -2.604358, -0.763921, 1.570796, 2.092951],accel_mss,speed_ms,0,blend_radius_m)
  movel([0.522304, -1.342219, -2.605587, -0.764582, 1.570796, 2.093101],accel_mss,speed_ms,0,blend_radius_m)
  movel([0.521907, -1.340536, -2.606678, -0.765175, 1.570796, 2.092703],accel_mss,speed_ms,0,blend_radius_m)
  movel([0.521520, -1.339809, -2.607147, -0.765432, 1.570796, 2.092316],accel_mss,speed_ms,0,blend_radius_m)
  speed_ms = 0.05
  movel([0.521520, -1.285564, -2.580155, -0.846670, 1.570796, 2.092316],accel_mss,speed_ms,0,blend_radius_m)
  speed_ms = 0.051
  movel([0.521520, -1.275543, -2.574496, -0.862350, 1.570796, 2.092316],accel_mss,speed_ms,0,blend_radius_m)
  movel([0.476022, -1.258693, -2.584253, -0.869443, 1.570796, 2.046818],accel_mss,speed_ms,0,blend_radius_m)
  movel([0.476022, -1.289833, -2.601246, -0.821310, 1.570796, 2.046818],accel_mss,speed_ms,0,blend_radius_m)
  speed_ms = 0.017
  movel([0.476022, -1.323578, -2.617448, -0.771363, 1.570796, 2.046818],accel_mss,speed_ms,0,blend_radius_m)
  speed_ms = 0.051
  movel([0.470953, -1.322609, -2.618052, -0.771728, 1.570796, 2.041749],accel_mss,speed_ms,0,blend_radius_m)
  movel([0.465499, -1.322151, -2.618337, -0.771902, 1.570796, 2.036295],accel_mss,speed_ms,0,blend_radius_m)
  movel([0.459700, -1.322218, -2.618295, -0.771876, 1.570796, 2.030497],accel_mss,speed_ms,0,blend_radius_m)
  movel([0.453607, -1.322817, -2.617922, -0.771650, 1.570796, 2.024404],accel_mss,speed_ms,0,blend_radius_m)
  movel([0.447278, -1.323954, -2.617214, -0.771222, 1.570796, 2.018074],accel_mss,speed_ms,0,blend_radius_m)
  movel([0.440789, -1.325614, -2.616175, -0.770599, 1.570796, 2.011585],accel_mss,speed_ms,0,blend_radius_m)
  movel([0.434220, -1.327782, -2.614814, -0.769792, 1.570796, 2.005017],accel_mss,speed_ms,0,blend_radius_m)
  movel([0.427664, -1.330421, -2.613149, -0.768819, 1.570796, 1.998461],accel_mss,speed_ms,0,blend_radius_m)
  movel([0.421211, -1.333492, -2.611199, -0.767698, 1.570796, 1.992008],accel_mss,speed_ms,0,blend_radius_m)
  movel([0.414946, -1.336944, -2.608992, -0.766453, 1.570796, 1.985742],accel_mss,speed_ms,0,blend_radius_m)
  movel([0.408955, -1.340716, -2.606561, -0.765112, 1.570796, 1.979752],accel_mss,speed_ms,0,blend_radius_m)
  movel([0.403302, -1.344754, -2.603937, -0.763697, 1.570796, 1.974099],accel_mss,speed_ms,0,blend_radius_m)
  movel([0.398041, -1.349002, -2.601153, -0.762234, 1.570796, 1.968837],accel_mss,speed_ms,0,blend_radius_m)
  movel([0.393215, -1.353405, -2.598240, -0.760743, 1.570796, 1.964011],accel_mss,speed_ms,0,blend_radius_m)
  movel([0.388847, -1.357921, -2.595225, -0.759243, 1.570796, 1.959643],accel_mss,speed_ms,0,blend_radius_m)
  movel([0.384950, -1.362513, -2.592130, -0.757747, 1.570796, 1.955746],accel_mss,speed_ms,0,blend_radius_m)
  movel([0.381534, -1.367152, -2.588972, -0.756265, 1.570796, 1.952330],accel_mss,speed_ms,0,blend_radius_m)
  movel([0.378599, -1.371819, -2.585764, -0.754806, 1.570796, 1.949395],accel_mss,speed_ms,0,blend_radius_m)
  movel([0.376141, -1.376502, -2.582514, -0.753373, 1.570796, 1.946938],accel_mss,speed_ms,0,blend_radius_m)
  movel([0.374160, -1.381191, -2.579228, -0.751970, 1.570796, 1.944957],accel_mss,speed_ms,0,blend_radius_m)
  movel([0.372653, -1.385882, -2.575909, -0.750598, 1.570796, 1.943450],accel_mss,speed_ms,0,blend_radius_m)
  movel([0.371623, -1.390576, -2.572555, -0.749258, 1.570796, 1.942419],accel_mss,speed_ms,0,blend_radius_m)
  movel([0.371073, -1.395273, -2.569167, -0.747948, 1.570796, 1.941869],accel_mss,speed_ms,0,blend_radius_m)
  movel([0.371012, -1.399975, -2.565744, -0.746670, 1.570796, 1.941809],accel_mss,speed_ms,0,blend_radius_m)
  movel([0.371456, -1.404683, -2.562282, -0.745423, 1.570796, 1.942252],accel_mss,speed_ms,0,blend_radius_m)
  movel([0.372418, -1.409403, -2.558780, -0.744206, 1.570796, 1.943215],accel_mss,speed_ms,0,blend_radius_m)
  movel([0.373917, -1.414134, -2.555236, -0.743019, 1.570796, 1.944713],accel_mss,speed_ms,0,blend_radius_m)
  movel([0.375977, -1.418879, -2.551647, -0.741863, 1.570796, 1.946774],accel_mss,speed_ms,0,blend_radius_m)
  movel([0.377107, -1.421048, -2.549995, -0.741346, 1.570796, 1.947904],accel_mss,speed_ms,0,blend_radius_m)
  movel([0.380371, -1.425022, -2.546951, -0.740416, 1.570796, 1.951168],accel_mss,speed_ms,0,blend_radius_m)
  movel([0.383894, -1.428548, -2.544229, -0.739611, 1.570796, 1.954690],accel_mss,speed_ms,0,blend_radius_m)
  movel([0.387547, -1.431518, -2.541923, -0.738948, 1.570796, 1.958343],accel_mss,speed_ms,0,blend_radius_m)
  movel([0.391324, -1.433965, -2.540012, -0.738412, 1.570796, 1.962120],accel_mss,speed_ms,0,blend_radius_m)
  movel([0.395214, -1.435924, -2.538476, -0.737989, 1.570796, 1.966011],accel_mss,speed_ms,0,blend_radius_m)
  movel([0.399213, -1.437422, -2.537297, -0.737670, 1.570796, 1.970009],accel_mss,speed_ms,0,blend_radius_m)
  movel([0.403317, -1.438485, -2.536458, -0.737446, 1.570796, 1.974113],accel_mss,speed_ms,0,blend_radius_m)
  movel([0.407527, -1.439130, -2.535949, -0.737310, 1.570796, 1.978323],accel_mss,speed_ms,0,blend_radius_m)
  movel([0.411841, -1.439371, -2.535758, -0.737260, 1.570796, 1.982637],accel_mss,speed_ms,0,blend_radius_m)
  movel([0.416265, -1.439219, -2.535879, -0.737292, 1.570796, 1.987061],accel_mss,speed_ms,0,blend_radius_m)
  movel([0.420797, -1.438676, -2.536308, -0.737405, 1.570796, 1.991594],accel_mss,speed_ms,0,blend_radius_m)
  movel([0.425441, -1.437743, -2.537044, -0.737602, 1.570796, 1.996238],accel_mss,speed_ms,0,blend_radius_m)
  movel([0.430197, -1.436417, -2.538088, -0.737884, 1.570796, 2.000993],accel_mss,speed_ms,0,blend_radius_m)
  movel([0.435055, -1.434695, -2.539440, -0.738254, 1.570796, 2.005852],accel_mss,speed_ms,0,blend_radius_m)
  movel([0.440009, -1.432571, -2.541102, -0.738716, 1.570796, 2.010806],accel_mss,speed_ms,0,blend_radius_m)
  movel([0.445042, -1.430040, -2.543073, -0.739277, 1.570796, 2.015839],accel_mss,speed_ms,0,blend_radius_m)
  movel([0.450131, -1.427099, -2.545350, -0.739940, 1.570796, 2.020927],accel_mss,speed_ms,0,blend_radius_m)
  movel([0.455238, -1.423758, -2.547922, -0.740709, 1.570796, 2.026035],accel_mss,speed_ms,0,blend_radius_m)
  movel([0.460327, -1.420025, -2.550776, -0.741589, 1.570796, 2.031124],accel_mss,speed_ms,0,blend_radius_m)
  movel([0.465347, -1.415920, -2.553889, -0.742580, 1.570796, 2.036144],accel_mss,speed_ms,0,blend_radius_m)
  movel([0.470239, -1.411475, -2.557232, -0.743682, 1.570796, 2.041035],accel_mss,speed_ms,0,blend_radius_m)
  movel([0.474941, -1.406731, -2.560767, -0.744891, 1.570796, 2.045738],accel_mss,speed_ms,0,blend_radius_m)
  movel([0.479393, -1.401738, -2.564452, -0.746199, 1.570796, 2.050190],accel_mss,speed_ms,0,blend_radius_m)
  movel([0.483535, -1.396550, -2.568241, -0.747598, 1.570796, 2.054331],accel_mss,speed_ms,0,blend_radius_m)
  movel([0.487309, -1.391227, -2.572088, -0.749074, 1.570796, 2.058105],accel_mss,speed_ms,0,blend_radius_m)
  movel([0.490667, -1.385828, -2.575947, -0.750614, 1.570796, 2.061464],accel_mss,speed_ms,0,blend_radius_m)
  movel([0.493579, -1.380405, -2.579781, -0.752203, 1.570796, 2.064375],accel_mss,speed_ms,0,blend_radius_m)
  movel([0.496011, -1.375013, -2.583551, -0.753826, 1.570796, 2.066807],accel_mss,speed_ms,0,blend_radius_m)
